// TwinCAT 3 PLC project _49001_01_BSM_762_V01_000_ISCOtherm
// libraries:
//   Tc2_EtherCAT, * (Beckhoff Automation GmbH)
//   Tc2_IoFunctions, * (Beckhoff Automation GmbH)
//   Tc2_Math, * (Beckhoff Automation GmbH)
//   Tc2_MC2, * (Beckhoff Automation GmbH)
//   Tc2_NC, * (Beckhoff Automation GmbH)
//   Tc2_NCI, * (Beckhoff Automation GmbH)
//   Tc2_SerialCom, * (Beckhoff Automation GmbH)
//   Tc2_Standard, * (Beckhoff Automation GmbH)
//   Tc2_System, * (Beckhoff Automation GmbH)
//   Tc2_Utilities, * (Beckhoff Automation GmbH)
//   Tc3_Module, * (Beckhoff Automation GmbH)
//   Lib1,1.0.0.0,riex
// project tree:
//   Data types/Machine/BECKHOFF/ ST_BECKHOFFDRIVETOPLC.TcDUT, ST_BECKHOFFDRIVE_REF.TcDUT, ST_PLCTOBECKHOFFDRIVE.TcDUT
//   Data types/Machine/FORCE/ ST_FORCETOPLC.TcDUT, ST_FORCE_REF.TcDUT, ST_PLCTOFORCE.TcDUT
//   Data types/Machine/Group_0000 - General/ ET_Gr00Auto.TcDUT, ET_Gr00Home.TcDUT, ST_Gr00HMIRef.TcDUT, ST_Gr00HMITOPLC.TcDUT, ST_Gr00PLCTOHMI.TcDUT
//   Data types/Machine/Group_0001/ ET_Gr01Auto.TcDUT, ET_Gr01Home.TcDUT, ET_Gr01HomeAxis.TcDUT, ET_Gr01HomeSawband.TcDUT, ET_Gr01Manual.TcDUT, ST_Gr01HMIRef.TcDUT, ST_Gr01HMITOPLC.TcDUT, ST_Gr01PLCTOHMI.TcDUT
//   Data types/Machine/Group_0002/ ET_Gr02Auto.TcDUT, ET_Gr02Home.TcDUT, ET_Gr02HomeAxis.TcDUT, ET_Gr02Manual.TcDUT, ST_Gr02HMIRef.TcDUT, ST_Gr02HMITOPLC.TcDUT, ST_Gr02PLCTOHMI.TcDUT
//   Data types/Machine/Group_0005/ ET_Gr05Auto.TcDUT, ET_Gr05AutoProcess.TcDUT, ET_Gr05Home.TcDUT, ET_Gr05HomeAxis.TcDUT, ET_Gr05HomeAxisClamp1.TcDUT, ET_Gr05Manual.TcDUT, ST_Gr05HMIRef.TcDUT, ST_Gr05HMITOPLC.TcDUT, ST_Gr05PLCTOHMI.TcDUT
//   Data types/Machine/SEW/CIA402/ ST_PLCTOSEWMOVIEDRIVEBCIA402.TcDUT, ST_SEWMOVIEDRIVEBCIA402TOPLC.TcDUT, ST_SEWMOVIEDRIVEBCIA402_REF.TcDUT
//   Data types/Machine/STOEBER/PS6A34/ ST_STOEBER_PS6A34Status.TcDUT
//   Data types/Machine/STOEBER/SDS/ ST_BaseDeviceIn.TcDUT, ST_BaseDeviceOut.TcDUT, ST_PLCTOSTOEBER.TcDUT, ST_STOEBERTOPLC.TcDUT
//   Data types/Machine/STOEBER/SI6_SC6/CIA402/ ST_CIA402In.TcDUT, ST_CIA402Out.TcDUT, ST_PLCTOSTOEBERSI6SC6CIA402.TcDUT, ST_STOEBERSI6SC6CIA402TOPLC.TcDUT, ST_STOEBERSI6SC6CIA402_REF.TcDUT
//   Data types/Machine/STOEBER/ ST_STOEBER_AxisStatus.TcDUT
//   Data types/Machine/WeldingPhases/ ET_WeldingDirection.TcDUT, ST_WeldingStatus.TcDUT
//   Data types/Machine/WeldingPhases/Force/ ST_BeadUp.TcDUT, ST_ForceProcess.TcDUT, ST_ForceWelding.TcDUT, ST_HeatUp.TcDUT, ST_PreHeat.TcDUT, ST_WeldingPhases.TcDUT
//   Data types/Machine/WeldingPhases/Position/ ST_PositionProcess.TcDUT, ST_PositionWelding.TcDUT
//   Data types/Objects/Axis/ExternelMC/ ET_JogMode.TcDUT, ET_MC_Direction.TcDUT, ET_MC_States.TcDUT, ST_AXIS_REF.TcDUT, ST_NCTOPLC.TcDUT, ST_PLCTONC.TcDUT
//   Data types/Objects/Axis/ExternelMC/SDS/ ST_CommandPositioningFROMNC.TcDUT, ST_CommandPositioningFROMPLC.TcDUT, ST_DRIVE_REF.TcDUT, ST_FastRefereneValueFROMNC.TcDUT, ST_FastRefereneValueFROMPLC.TcDUT
//   Data types/Objects/Axis/ExternelMC/SI6/ ET_ModesOfOperation.TcDUT, ST_DRIVESI6SC6CIA402_REF.TcDUT, ST_HomingModeFromDrive.TcDUT, ST_HomingModeFromPLC.TcDUT, ST_JogModeFromPLC.TcDUT, ST_PositionModeFromDrive.TcDUT, ST_PositionModeFromPLC.TcDUT, ST_TorqueModeFromDrive.TcDUT, ST_TorqueModeFromPLC.TcDUT, ST_VelocityModeFromDrive.TcDUT, ST_VelocityModeFromPLC.TcDUT
//   Data types/Objects/Axis/InternalMC/Controller/ ET_MC_ControllerMode.TcDUT, ST_VeloControllerConfig.TcDUT
//   Data types/Objects/Axis/InternalMC/Drive/Control/ ST_AxisCtrl.TcDUT (not stored), ST_TippingMode.TcDUT (not stored)
//   Data types/Objects/Axis/InternalMC/Drive/Parameter/ ST_Dynamics.TcDUT (not stored), ST_LimitSwitches.TcDUT (not stored), ST_Position.TcDUT (not stored)
//   Data types/Objects/Axis/InternalMC/Drive/Scaling/ ET_MC_RampType.TcDUT (not stored), ET_ScalingMethod.TcDUT (not stored), ST_Scaling.TcDUT (not stored)
//   Data types/Objects/Axis/InternalMC/Drive/States/ ET_MC_MotionStates.TcDUT (not stored), ST_AxisStates.TcDUT (not stored)
//   Data types/Objects/Axis/InternalMC/Drive/ ST_DriveConfig.TcDUT
//   Data types/Objects/Axis/InternalMC/Encoder/ ST_EncoderConfig.TcDUT
//   Data types/Objects/Axis/InternalMC/ ST_AXIS_REF_V2.TcDUT
//   Data types/Objects/EtherCAT Diag/ ET_EtherCATDiag.TcDUT, E_EcCommState.TcDUT, ST_EcMasterDevState.TcDUT, ST_SlaveState.TcDUT, ST_SlaveStateInfo.TcDUT, ST_SlaveStateInfoScanned.TcDUT, ST_TopologyData.TcDUT
//   Data types/Objects/ET_SpindleCtrl/ ET_SpindleCtrl.TcDUT
//   Data types/Objects/FB_Alarm/ ET_AlarmType.TcDUT, ST_Alarm.TcDUT, ST_AlarmIn.TcDUT, ST_AlarmOut.TcDUT, ST_AlarmProperties.TcDUT, ST_AlarmRef.TcDUT
//   Data types/Objects/FB_AxisController/ ET_AxisGetLimits.TcDUT, ET_AxisSetLimits.TcDUT, ET_STOEBER_AxisGetLimitsTc2.TcDUT, ET_STOEBER_AxisSetLimitsTc2.TcDUT
//   Data types/Objects/FB_AxisMoveManual/ ET_AxisMoveManualSetLimits.TcDUT
//   Data types/Objects/FB_Blinker/ ST_Blinker.TcDUT
//   Data types/Objects/FB_CalcContour/ ET_ContourType.TcDUT
//   Data types/Objects/FB_CfgAxisInExt3DGroup/ ET_CfgAxisInExt3DGroup.TcDUT
//   Data types/Objects/FB_DistanceCounter/ ST_DistanceCounter.TcDUT
//   Data types/Objects/FB_EL3312/ ET_EL3312ThermocoupleTyp.TcDUT, ST_EL3312ChannelState.TcDUT, ST_EL3312CoeInfo.TcDUT, ST_EL3312CoeReadData.TcDUT, ST_EL3312CoeWriteData.TcDUT
//   Data types/Objects/FB_EL3351/ ST_EL3351ChannelState.TcDUT, ST_EL3351CoeInfo.TcDUT, ST_EL3351CoeReadData.TcDUT, ST_EL3351CoeWriteData.TcDUT
//   Data types/Objects/FB_EL3356/ ST_EL3356ChannelCtrl.TcDUT, ST_EL3356ChannelState.TcDUT, ST_EL3356CoeInfo.TcDUT, ST_EL3356CoeReadData.TcDUT, ST_EL3356CoeWriteData.TcDUT
//   Data types/Objects/FB_ExtSetPoint/ ET_MoveExtState.TcDUT
//   Data types/Objects/FB_ExtTrajPos/ ET_CalcExtTrajState.TcDUT
//   Data types/Objects/FB_ItpReadRParams/ ET_ItpReadRParams.TcDUT
//   Data types/Objects/FB_ItpWriteRParams/ ET_ItpWriteRParams.TcDUT
//   Data types/Objects/FB_KL600x/ ET_KL600xInit.TcDUT, ET_KL600xSend.TcDUT, ST_KL600xData.TcDUT
//   Data types/Objects/FB_LoadFromFile/ ET_LoadFromFile.TcDUT
//   Data types/Objects/FB_Logger/ ST_Logger.TcDUT, ST_LoggerVar.TcDUT
//   Data types/Objects/FB_ModeSelector/ ET_MachineMode.TcDUT, ET_MachineState.TcDUT
//   Data types/Objects/FB_RampDirector/ ET_RampGenerator.TcDUT
//   Data types/Objects/FB_SpindlePreheat/ ET_SpindlePreheat.TcDUT, ST_SpindlePreheat.TcDUT
//   Data types/Objects/FB_TimeHoursCounter/ ST_TimeHoursCounter.TcDUT
//   Data types/Objects/FB_Timer/ ST_DateTime.TcDUT, ST_Time.TcDUT
//   Data types/Objects/FB_ToolStorage/ ET_ToolStatus.TcDUT, ET_ToolStorage.TcDUT
//   Data types/Objects/FB_Traceability/ ST_Traceability.TcDUT, ST_TraceabilityData.TcDUT, ST_TraceabilitySettings.TcDUT
//   Data types/Objects/Fieldbus/ ST_FieldbusStatus.TcDUT
//   Data types/Objects/Gefran/ ET_GFX4IR.TcDUT, ST_GFX4IRTOPLC.TcDUT, ST_GFX4IR_REF.TcDUT, ST_PLCTOGFX4IR.TcDUT
//   Data types/Objects/Leister/ ET_LeisterExtruder.TcDUT, ET_LeisterHeater.TcDUT, ST_LEISTERTOPLC.TcDUT, ST_LEISTER_REF.TcDUT, ST_PLCTOLEISTER.TcDUT
//   Data types/Objects/Munsch/ ET_MunschExtruder.TcDUT, ET_MUNSCH_CMD.TcDUT, ET_MUNSCH_RES.TcDUT, ST_MUNSCH_CMD_Data.TcDUT, ST_MUNSCH_REF.TcDUT, ST_MUNSCH_RES_Data.TcDUT
//   Data types/Objects/Periphery/ ST_PERIPHERYTOPLC.TcDUT, ST_PERIPHERY_REF.TcDUT, ST_PLCTOPERIPHERY.TcDUT
//   Data types/Objects/Robot/KUKA/ ET_KukaStart.TcDUT, ST_KUKATOPLC.TcDUT, ST_KUKA_REF.TcDUT, ST_PLCTOKUKA.TcDUT
//   Data types/Objects/Robot/ ST_PLCTOROBOT.TcDUT, ST_ROBOTTOPLC.TcDUT
//   Data types/Objects/Robot/YASKAWA/ ET_YaskawaStart.TcDUT, ST_PLCTOYASKAWA.TcDUT, ST_YASKAWATOPLC.TcDUT, ST_YASKAWA_REF.TcDUT
//   Data types/Objects/Spindle/ ET_SpindleClutchStatus.TcDUT
//   Data types/Objects/Spindle/PDS/ ST_SpindlePDSXLA170ClutchStatus.TcDUT, ST_SpindlePDSXLHClutchStatus.TcDUT
//   Data types/Objects/Terminal/ ST_TerminalState.TcDUT
//   Data types/Objects/TouchProbe/Renishaw/ ST_TouchProbeRenishawCtrl.TcDUT, ST_TouchProbeRenishawStatus.TcDUT
//   Data types/Objects/VFD/ ST_PLCTOVFD.TcDUT, ST_VFDTOPLC.TcDUT, ST_VFD_AXIS_REF.TcDUT, ST_VFD_DRIVE_REF.TcDUT
//   Global Variables/Alarms/ GVL_Gr00Alarm.TcGVL, GVL_Gr01Alarm.TcGVL, GVL_Gr02Alarm.TcGVL, GVL_Gr05Alarm.TcGVL
//   Global Variables/Basics/ GVL_FB_CheckArrayBounds.TcGVL, GVL_FB_CheckDivRealInfo.TcGVL
//   Global Variables/Config/ GVL_Gr00Config.TcGVL, GVL_Gr01Config.TcGVL, GVL_Gr02Config.TcGVL, GVL_Gr05Config.TcGVL
//   Global Variables/FB_Alarm/ GVL_FB_Alarm.TcGVL
//   Global Variables/FB_Fieldbus/ GVL_FB_Fieldbus.TcGVL
//   Global Variables/FB_GFX4IRZones/ GVL_FB_GFX4IRZones.TcGVL
//   Global Variables/FB_LoadFromFile/ GVL_FB_LoadFromFile.TcGVL
//   Global Variables/FB_Logger/ GVL_FB_Logger.TcGVL
//   Global Variables/FB_Traceability/ GVL_Traceability.TcGVL
//   Global Variables/ GVL.TcGVL, GVL_Gr0000.TcGVL, GVL_Gr0100.TcGVL, GVL_Gr0200.TcGVL, GVL_Gr0500.TcGVL, TwinCAT_Import.TcGVL
//   Global Variables/HMI/ GVL_Gr00HMI.TcGVL, GVL_Gr01HMI.TcGVL, GVL_Gr02HMI.TcGVL, GVL_Gr05HMI.TcGVL
//   Global Variables/Init/ GVL_Gr00Init.TcGVL, GVL_Gr01Init.TcGVL, GVL_Gr02Init.TcGVL, GVL_Gr05Init.TcGVL
//   Global Variables/Interface/ GVL_Gr00Interface.TcGVL, GVL_Gr01Interface.TcGVL, GVL_Gr02Interface.TcGVL, GVL_Gr05Interface.TcGVL
//   Global Variables/IO/ GVL_Gr00IO.TcGVL, GVL_Gr01IO.TcGVL, GVL_Gr02IO.TcGVL, GVL_Gr05IO.TcGVL
//   / PLC_TASK.TcTTO, Recipe Manager.TcRMO (not stored) (excluded from build)
//   POUs/ FAST.TcPOU, Init.TcPOU, MAIN.TcPOU
//   POUs/Machine/Group_0000 - General/Gr00Alarm/ FB_Gr00Alarm.TcPOU
//   POUs/Machine/Group_0000 - General/Gr00Control/ Gr00Control.TcPOU
//   POUs/Machine/Group_0000 - General/Gr00Control/Gr00Periphery/ FB_Gr00Periphery.TcPOU
//   POUs/Machine/Group_0000 - General/Gr00Control/Gr00Program/ FB_Gr00Program.TcPOU
//   POUs/Machine/Group_0000 - General/Gr00Control/Gr00Safety/ FB_Gr00Safety.TcPOU
//   POUs/Machine/Group_0000 - General/Gr00Control/Gr00Signals/ FB_Gr00Signals.TcPOU
//   POUs/Machine/Group_0000 - General/Gr00Control/Gr00Utility/ FB_Gr00Utility.TcPOU
//   POUs/Machine/Group_0000 - General/ Gr00Coordinator.TcPOU
//   POUs/Machine/Group_0000 - General/Gr00MachineMode/Gr00Auto/ Gr00Auto.TcPOU
//   POUs/Machine/Group_0000 - General/Gr00MachineMode/Gr00Auto/Gr00AutoAlarm/ FB_Gr00AutoAlarm.TcPOU (not stored)
//   POUs/Machine/Group_0000 - General/Gr00MachineMode/Gr00Auto/Gr00AutoInit/ FB_Gr00AutoInit.TcPOU (not stored)
//   POUs/Machine/Group_0000 - General/Gr00MachineMode/Gr00Auto/Gr00AutoProcedure/ FB_Gr00AutoProcedure.TcPOU (not stored)
//   POUs/Machine/Group_0000 - General/Gr00MachineMode/Gr00HMI/ Gr00HMI.TcPOU
//   POUs/Machine/Group_0000 - General/Gr00MachineMode/Gr00Home/ Gr00Home.TcPOU
//   POUs/Machine/Group_0000 - General/Gr00MachineMode/Gr00Home/Gr00HomeAlarm/ FB_Gr00HomeAlarm.TcPOU (not stored)
//   POUs/Machine/Group_0000 - General/Gr00MachineMode/Gr00Home/Gr00HomeInit/ FB_Gr00HomeInit.TcPOU (not stored)
//   POUs/Machine/Group_0000 - General/Gr00MachineMode/Gr00Home/Gr00HomeProcedure/ FB_Gr00HomeProcedure.TcPOU (not stored)
//   POUs/Machine/Group_0000 - General/Gr00MachineMode/ Gr00MachineMode.TcPOU
//   POUs/Machine/Group_0000 - General/Gr00MachineMode/Gr00Manual/ Gr00Manual.TcPOU
//   POUs/Machine/Group_0000 - General/Gr00MachineMode/Gr00Manual/Gr00ManualAlarm/ FB_Gr00ManualAlarm.TcPOU (not stored)
//   POUs/Machine/Group_0000 - General/Gr00MachineMode/Gr00Manual/Gr00ManualInit/ FB_Gr00ManualInit.TcPOU (not stored)
//   POUs/Machine/Group_0000 - General/Gr00MachineMode/Gr00Manual/Gr00ManualProcedure/ FB_Gr00ManualProcedure.TcPOU (not stored)
//   POUs/Machine/Group_0000 - General/Gr00Persistent/ Gr00Persistent.TcPOU
//   POUs/Machine/Group_0000 - General/Gr00Simulation/ Gr00Simulation.TcPOU
//   POUs/Machine/Group_0100 - Production/Gr01Control/Gr01Alarm/ FB_Gr01Alarm.TcPOU
//   POUs/Machine/Group_0100 - Production/Gr01Control/ Gr01Control.TcPOU
//   POUs/Machine/Group_0100 - Production/Gr01Control/Gr01Safety/ FB_Gr01Safety.TcPOU
//   POUs/Machine/Group_0100 - Production/Gr01Control/Gr01Signals/ FB_Gr01Signals.TcPOU
//   POUs/Machine/Group_0100 - Production/Gr01Control/Gr01Units/ FB_Gr01Angle.TcPOU, FB_Gr01SawBow.TcPOU
//   POUs/Machine/Group_0100 - Production/Gr01Control/Gr01Units/FB_Gr01Sawband/ FB_Gr01Sawband.TcPOU (not stored), FB_LowPassFilter.TcPOU (not stored), FB_PosVeloEnc.TcPOU (not stored)
//   POUs/Machine/Group_0100 - Production/Gr01Control/Gr01Utility/ FB_Gr01Utility.TcPOU
//   POUs/Machine/Group_0100 - Production/ Gr01Coordinator.TcPOU
//   POUs/Machine/Group_0100 - Production/Gr01HMI/ Gr01HMI.TcPOU
//   POUs/Machine/Group_0100 - Production/Gr01MachineMode/Gr01Auto/ Gr01Auto.TcPOU
//   POUs/Machine/Group_0100 - Production/Gr01MachineMode/Gr01Auto/Gr01AutoAlarm/ FB_Gr01AutoAlarm.TcPOU (not stored)
//   POUs/Machine/Group_0100 - Production/Gr01MachineMode/Gr01Auto/Gr01AutoInit/ FB_Gr01AutoInit.TcPOU (not stored)
//   POUs/Machine/Group_0100 - Production/Gr01MachineMode/Gr01Auto/Gr01AutoProcedure/ FB_Gr01AutoProcedure.TcPOU (not stored)
//   POUs/Machine/Group_0100 - Production/Gr01MachineMode/Gr01Home/ Gr01Home.TcPOU
//   POUs/Machine/Group_0100 - Production/Gr01MachineMode/Gr01Home/Gr01HomeAlarm/ FB_Gr01HomeAlarm.TcPOU (not stored)
//   POUs/Machine/Group_0100 - Production/Gr01MachineMode/Gr01Home/Gr01HomeFunctions/ FB_Gr01HomeAngle.TcPOU (not stored), FB_Gr01HomeAxisSawBow.TcPOU (not stored), FB_Gr01HomeSawband.TcPOU (not stored)
//   POUs/Machine/Group_0100 - Production/Gr01MachineMode/Gr01Home/Gr01HomeInit/ FB_Gr01HomeInit.TcPOU (not stored)
//   POUs/Machine/Group_0100 - Production/Gr01MachineMode/Gr01Home/Gr01HomeProcedure/ FB_Gr01HomeProcedure.TcPOU (not stored)
//   POUs/Machine/Group_0100 - Production/Gr01MachineMode/ Gr01MachineMode.TcPOU
//   POUs/Machine/Group_0100 - Production/Gr01MachineMode/Gr01Manual/ Gr01Manual.TcPOU
//   POUs/Machine/Group_0100 - Production/Gr01MachineMode/Gr01Manual/Gr01ManualAlarm/ FB_Gr01ManualAlarm.TcPOU (not stored)
//   POUs/Machine/Group_0100 - Production/Gr01MachineMode/Gr01Manual/Gr01ManualInit/ FB_Gr01ManualInit.TcPOU (not stored)
//   POUs/Machine/Group_0100 - Production/Gr01MachineMode/Gr01Manual/Gr01ManualProcedure/ FB_Gr01ManualProcedure.TcPOU (not stored)
//   POUs/Machine/Group_0100 - Production/Gr01Persistent/ Gr01Persistent.TcPOU
//   POUs/Machine/Group_0100 - Production/Gr01Simulation/ Gr01Simulation.TcPOU
//   POUs/Machine/Group_0500 - Transport/Gr05Control/Gr05Alarm/ FB_Gr05Alarm.TcPOU
//   POUs/Machine/Group_0500 - Transport/Gr05Control/ Gr05Control.TcPOU
//   POUs/Machine/Group_0500 - Transport/Gr05Control/Gr05Safety/ FB_Gr05Safety.TcPOU
//   POUs/Machine/Group_0500 - Transport/Gr05Control/Gr05Signals/ FB_Gr05Signals.TcPOU
//   POUs/Machine/Group_0500 - Transport/Gr05Control/Gr05Units/ FB_Gr05AxisClamp.TcPOU, FB_Gr05CylinderClamp.TcPOU, FB_Gr05CylinderPos.TcPOU, FB_Gr05RemovalBand.TcPOU, FB_Gr05Slide.TcPOU
//   POUs/Machine/Group_0500 - Transport/Gr05Control/Gr05Utility/ FB_Gr05Utility.TcPOU
//   POUs/Machine/Group_0500 - Transport/ Gr05Coordinator.TcPOU
//   POUs/Machine/Group_0500 - Transport/Gr05HMI/ Gr05HMI.TcPOU
//   POUs/Machine/Group_0500 - Transport/Gr05MachineMode/Gr05Auto/ Gr05Auto.TcPOU
//   POUs/Machine/Group_0500 - Transport/Gr05MachineMode/Gr05Auto/Gr05AutoAlarm/ FB_Gr05AutoAlarm.TcPOU (not stored)
//   POUs/Machine/Group_0500 - Transport/Gr05MachineMode/Gr05Auto/Gr05AutoInit/ FB_Gr05AutoInit.TcPOU (not stored)
//   POUs/Machine/Group_0500 - Transport/Gr05MachineMode/Gr05Auto/Gr05AutoProcedure/ FB_Gr05AutoProcedure.TcPOU (not stored)
//   POUs/Machine/Group_0500 - Transport/Gr05MachineMode/Gr05Home/ Gr05Home.TcPOU
//   POUs/Machine/Group_0500 - Transport/Gr05MachineMode/Gr05Home/Gr05HomeAlarm/ FB_Gr05HomeAlarm.TcPOU (not stored)
//   POUs/Machine/Group_0500 - Transport/Gr05MachineMode/Gr05Home/Gr05HomeFunctions/ FB_Gr05HomeAxisClamp1.TcPOU (not stored), FB_Gr05HomeAxisClamp2.TcPOU (not stored)
//   POUs/Machine/Group_0500 - Transport/Gr05MachineMode/Gr05Home/Gr05HomeInit/ FB_Gr05HomeInit.TcPOU (not stored)
//   POUs/Machine/Group_0500 - Transport/Gr05MachineMode/Gr05Home/Gr05HomeProcedure/ FB_Gr05HomeProcedure.TcPOU (not stored)
//   POUs/Machine/Group_0500 - Transport/Gr05MachineMode/ Gr05MachineMode.TcPOU
//   POUs/Machine/Group_0500 - Transport/Gr05MachineMode/Gr05Manual/ Gr05Manual.TcPOU
//   POUs/Machine/Group_0500 - Transport/Gr05MachineMode/Gr05Manual/Gr05ManualAlarm/ FB_Gr05ManualAlarm.TcPOU (not stored)
//   POUs/Machine/Group_0500 - Transport/Gr05MachineMode/Gr05Manual/Gr05ManualInit/ FB_Gr05ManualInit.TcPOU (not stored)
//   POUs/Machine/Group_0500 - Transport/Gr05MachineMode/Gr05Manual/Gr05ManualProcedure/ FB_Gr05ManualProcedure.TcPOU (not stored)
//   POUs/Machine/Group_0500 - Transport/Gr05Persistent/ Gr05Persistent.TcPOU
//   POUs/Machine/Group_0500 - Transport/Gr05Simulation/ Gr05Simulation.TcPOU
//   POUs/Tc2 Objects/Alarm/ FB_Alarm.TcPOU, FB_Error.TcPOU, FB_FatalError.TcPOU, FB_Hint.TcPOU, FB_Message.TcPOU, FB_Warning.TcPOU
//   POUs/Tc2 Objects/Automation/Axis/Beckhoff/CommandPositioning/ FB_AxisController.TcPOU (not stored), FB_AxisMoveAuto.TcPOU (not stored), FB_AxisMoveManual.TcPOU (not stored)
//   POUs/Tc2 Objects/Automation/Axis/Beckhoff/ FB_AxisMcBeckhoff.TcPOU, FB_AxisMcBeckhoffSEWMoviDriveBVelo.TcPOU, FB_AxisMcBeckhoffStoeberSCI6.TcPOU, FB_BECKHOFFDRIVE_REF.TcPOU
//   POUs/Tc2 Objects/Automation/Axis/ F_ChkAllAxisCoupled.TcPOU, F_ChkAllAxisEnabled.TcPOU, F_ChkAllAxisFieldbusOK.TcPOU, F_ChkAllAxisInSamePos.TcPOU, F_ChkAllAxisNotMoving.TcPOU, F_ChkAllAxisReferenced.TcPOU, F_ChkAllAxisStandStill.TcPOU
//   POUs/Tc2 Objects/Automation/Axis/OnOff/ FB_OnOff_AxisController.TcPOU, FB_OnOff_AxisMoveAuto.TcPOU, FB_OnOff_AxisMoveManual.TcPOU
//   POUs/Tc2 Objects/Automation/Axis/OnOff/Motion/ FB_OnOff_MoveAbsolut.TcPOU (not stored), FB_OnOff_MoveVelocity.TcPOU (not stored), FB_OnOff_Power.TcPOU (not stored), FB_OnOff_Reset.TcPOU (not stored), FB_OnOff_Stop.TcPOU (not stored)
//   POUs/Tc2 Objects/Automation/Axis/Override/ FB_Override.TcPOU, FB_OverrideSelection.TcPOU
//   POUs/Tc2 Objects/Automation/Axis/Own/Interface/Drive/ FB_AXIS_REF_V2.TcPOU (not stored)
//   POUs/Tc2 Objects/Automation/Axis/SEW/MOVIDRIVE B/ FB_SEWMOVIDRIVEBCIA402_REF.TcPOU (not stored)
//   POUs/Tc2 Objects/Automation/Axis/Stöber/SDS/CommandPositioning/ FB_AxisMcStoeber.TcPOU (not stored), FB_STOEBERSDS_MC_AxisController.TcPOU (not stored), FB_STOEBERSDS_MC_AxisMoveAuto.TcPOU (not stored), FB_STOEBERSDS_MC_AxisMoveManual.TcPOU (not stored), FB_STOEBERSDS_MC_GearIn.TcPOU (not stored), FB_STOEBERSDS_MC_GearOut.TcPOU (not stored), FB_STOEBERSDS_MC_Halt_noready.TcPOU (not stored), FB_STOEBERSDS_MC_Home.TcPOU (not stored), FB_STOEBERSDS_MC_Jog.TcPOU (not stored), FB_STOEBERSDS_MC_MoveAbsolut.TcPOU (not stored), FB_STOEBERSDS_MC_MoveAdditive.TcPOU (not stored), FB_STOEBERSDS_MC_MoveRelative.TcPOU (not stored), FB_STOEBERSDS_MC_MoveSuperimposed.TcPOU (not stored), FB_STOEBERSDS_MC_MoveVelocity.TcPOU (not stored), FB_STOEBERSDS_MC_Power.TcPOU (not stored), FB_STOEBERSDS_MC_Reset.TcPOU (not stored), FB_STOEBERSDS_MC_Stop.TcPOU (not stored), F_MoveToAxisRef.TcPOU (not stored)
//   POUs/Tc2 Objects/Automation/Axis/Stöber/SDS/FastRefereneValue/ FB_AxisStoeberSDS.TcPOU (not stored), FB_STOEBERSDS_AxisController.TcPOU (not stored), FB_STOEBERSDS_AxisMoveAuto.TcPOU (not stored), FB_STOEBERSDS_AxisMoveManual.TcPOU (not stored), FB_STOEBERSDS_Drive_REF.TcPOU (not stored), FB_STOEBERSDS_Home.TcPOU (not stored), FB_STOEBERSDS_Jog.TcPOU (not stored), FB_STOEBERSDS_MoveAbsolut.TcPOU (not stored), FB_STOEBERSDS_MoveVelocity.TcPOU (not stored), FB_STOEBERSDS_Power.TcPOU (not stored), FB_STOEBERSDS_QuickStop.TcPOU (not stored), FB_STOEBERSDS_Reset.TcPOU (not stored), FB_STOEBERSDS_Stop.TcPOU (not stored)
//   POUs/Tc2 Objects/Automation/Axis/Stöber/SDS/ FB_STOEBERSDS_AxisLink.TcPOU (not stored), FB_STOEBERSDS_ReadStatus.TcPOU (not stored)
//   POUs/Tc2 Objects/Automation/Axis/Stöber/SI6_SC6/ FB_StoeberPS6A34.TcPOU (not stored)
//   POUs/Tc2 Objects/Automation/Axis/VFD/ FB_VFD_AxisController.TcPOU, FB_VFD_AxisLink.TcPOU, FB_VFD_AxisMoveAuto.TcPOU, FB_VFD_AxisMoveManual.TcPOU (not stored), FB_VFD_Axis_REF.TcPOU (not stored), FB_VFD_Drive_REF.TcPOU (not stored), FB_VFD_MoveVelocity.TcPOU (not stored), FB_VFD_Power.TcPOU (not stored), FB_VFD_Reset.TcPOU (not stored), FB_VFD_Stop.TcPOU (not stored)
//   POUs/Tc2 Objects/Automation/Cylinder/ FB_Cylinder.TcPOU
//   POUs/Tc2 Objects/Automation/Cylinder/Hydraulic/ FB_HydraulicCylinder.TcPOU (not stored)
//   POUs/Tc2 Objects/Automation/Cylinder/Pneumatic/ FB_PneumaticCylinder.TcPOU (not stored)
//   POUs/Tc2 Objects/Automation/Cylinder/Position Cylinder/ FB_CylinderPos.TcPOU (not stored), FB_CylinderPos_MoveAbsolut.TcPOU (not stored), F_GetCylinderPos.TcPOU (not stored), F_SetCylinderPos.TcPOU (not stored)
//   POUs/Tc2 Objects/Automation/Extraction Fan/ FB_ExtractionFan.TcPOU
//   POUs/Tc2 Objects/Automation/Force/ FB_ForceController.TcPOU, FB_ForceReg.TcPOU, FB_FORCE_REF.TcPOU, FB_PID_Regler.TcPOU
//   POUs/Tc2 Objects/Automation/Heater/ FB_Heater.TcPOU
//   POUs/Tc2 Objects/Automation/MotorOnOff/ FB_Motor.TcPOU
//   POUs/Tc2 Objects/Automation/NCiChannel/ FB_CfgAxisInExt3DGroup.TcPOU
//   POUs/Tc2 Objects/Automation/NCiChannel/R-parameters/ FB_ItpReadRParams.TcPOU (not stored), FB_ItpWriteRParams.TcPOU (not stored)
//   POUs/Tc2 Objects/Automation/OperationMode/ FB_ModeSelector.TcPOU
//   POUs/Tc2 Objects/Automation/Process/ FB_StartProcess.TcPOU
//   POUs/Tc2 Objects/Automation/Sawband/ FB_Sawband.TcPOU
//   POUs/Tc2 Objects/Automation/Spindle/ FB_CoolingDevice.TcPOU, FB_SpindlePreheat.TcPOU, FB_ToolStorage.TcPOU, FB_VFD_SpindlePreheat.TcPOU, F_SpindleHSDClutchStatus.TcPOU, F_SpindlePDSXLA170ClutchStatus.TcPOU, F_SpindlePDSXLHClutchStatus.TcPOU
//   POUs/Tc2 Objects/Automation/Vacuum/ FB_Vacuum.TcPOU
//   POUs/Tc2 Objects/Basics/ CheckBounds.TcPOU (excluded from build), CheckDivReal.TcPOU (excluded from build), FB_CheckArrayBounds.TcPOU (excluded from build), FB_CheckDivRealInfo.TcPOU (excluded from build), FB_Get_Time.TcPOU, F_AdsError_Text.TcPOU
//   POUs/Tc2 Objects/Conversions/BitOriented/ F_ConvArrBitsToWord.TcPOU
//   POUs/Tc2 Objects/Diagnostic/Terminal/ FB_TerminalDiagnosis.TcPOU, FB_ToggleBit.TcPOU, F_StateReturn.TcPOU
//   POUs/Tc2 Objects/Engineering/Buffer/ FB_FiFo.TcPOU
//   POUs/Tc2 Objects/Engineering/Dynamics/CalcVeloAccDecJerk/ FB_CalcVeloAccDecJerk.TcPOU (not stored)
//   POUs/Tc2 Objects/Engineering/External set value generator/ FB_ExtSetPoint.TcPOU
//   POUs/Tc2 Objects/Engineering/Filter/ FB_PT1.TcPOU, FB_ValueFilter.TcPOU
//   POUs/Tc2 Objects/Engineering/Position offset/ F_PosOffset.TcPOU
//   POUs/Tc2 Objects/Engineering/Position/Controller/PID Components/ FB_CompD.TcPOU (not stored), FB_CompI.TcPOU (not stored), FB_CompP.TcPOU (not stored)
//   POUs/Tc2 Objects/Engineering/Position/Controller/PID Controller/ FB_CtrlOut.TcPOU (not stored), FB_CtrlPI.TcPOU (not stored), FB_CtrlPID.TcPOU (not stored), F_CtrlIn.TcPOU (not stored)
//   POUs/Tc2 Objects/Engineering/Position/Controller/PID Types/ FB_TypePI.TcPOU (not stored), FB_TypePID.TcPOU (not stored), FB_TypePIDW.TcPOU (not stored), FB_TypePIW.TcPOU (not stored)
//   POUs/Tc2 Objects/Engineering/Position/Controller/PositionController/ FB_PosCtrlIn.TcPOU (not stored), FB_PosCtrlOut.TcPOU (not stored), FB_PositionController.TcPOU (not stored)
//   POUs/Tc2 Objects/Engineering/Position/Encoder/ FB_PositionEncoder.TcPOU (not stored)
//   POUs/Tc2 Objects/Engineering/Position/ F_ModuloDistance.TcPOU
//   POUs/Tc2 Objects/Engineering/Position/Residuals/ F_ConvertActPosResiduals.TcPOU (not stored), F_ConvertSetPosResiduals.TcPOU (not stored)
//   POUs/Tc2 Objects/Engineering/Trajectory model/ FB_ExtContour.TcPOU, FB_ExtTraj.TcPOU, F_CalcContour.TcPOU, F_CalcTrajPos.TcPOU
//   POUs/Tc2 Objects/ExternalHardware/Beckhoff/EL..KL600x/ FB_KL600xData.TcPOU (not stored), FB_KL600xString.TcPOU (not stored)
//   POUs/Tc2 Objects/ExternalHardware/Beckhoff/EL3312/ FB_EL3312.TcPOU (not stored), FB_EL3312ChannelDiagnosis.TcPOU (not stored), FB_EL3312CoE.TcPOU (not stored)
//   POUs/Tc2 Objects/ExternalHardware/Beckhoff/EL3351/ FB_EL3351.TcPOU (not stored), FB_EL3351ChannelDiagnosis.TcPOU (not stored), FB_EL3351CoE.TcPOU (not stored), FB_EL3351Measuring.TcPOU (not stored)
//   POUs/Tc2 Objects/ExternalHardware/Beckhoff/EL3356/ FB_EL3356.TcPOU (not stored), FB_EL3356ChannelDiagnosis.TcPOU (not stored), FB_EL3356CoE.TcPOU (not stored)
//   POUs/Tc2 Objects/ExternalHardware/Gefran/ FB_GFX4IRCtrlZone.TcPOU, FB_GFX4IRZones.TcPOU, FB_GFX4IR_REF.TcPOU, F_ChkAllZonesNotEnabled.TcPOU
//   POUs/Tc2 Objects/ExternalHardware/KUKA/ FB_KUKA_Enable.TcPOU, FB_KUKA_Power.TcPOU, FB_KUKA_Prg.TcPOU, FB_KUKA_REF.TcPOU, FB_KUKA_Reset.TcPOU, FB_KUKA_StartProg.TcPOU, FB_MoveToKukaRef.TcPOU
//   POUs/Tc2 Objects/ExternalHardware/Leister/ FB_LeisterExtruder_Extruder.TcPOU, FB_LeisterExtruder_Heater.TcPOU, FB_LEISTER_EXTRUDER_REF.TcPOU
//   POUs/Tc2 Objects/ExternalHardware/Munsch/ FB_MunschExtruder.TcPOU, FB_MunschExtruderAir.TcPOU, FB_MunschExtruder_AirTemp.TcPOU, FB_MunschExtruder_Extruding.TcPOU, FB_MunschExtruder_Heat.TcPOU, FB_MunschExtruder_MaterialTemp.TcPOU, FB_MunschExtruder_ReadStatus.TcPOU, FB_MUNSCH_EXTRUDER_REF.TcPOU, F_MunschCMD.TcPOU, F_MunschRES.TcPOU
//   POUs/Tc2 Objects/ExternalHardware/Periphery/ FB_PERIPHERY_REF.TcPOU
//   POUs/Tc2 Objects/ExternalHardware/YASKAWA/ FB_YASKAWA_Controller.TcPOU, FB_YASKAWA_Power.TcPOU, FB_YASKAWA_REF.TcPOU, FB_YASKAWA_Reset.TcPOU, FB_YASKAWA_StartPrg.TcPOU
//   POUs/Tc2 Objects/File/ FB_FileHandler.TcPOU, FB_FileHandlerBinary.TcPOU, FB_LoadFromFile.TcPOU
//   POUs/Tc2 Objects/Logger/ FB_Logger.TcPOU, FB_LoggerFile.TcPOU
//   POUs/Tc2 Objects/Logic/ F_DwordToBitReal.TcPOU, F_RealToBitDword.TcPOU, F_ResetBitOfDWord.TcPOU, F_SetBitOfDWord.TcPOU
//   POUs/Tc2 Objects/Logic/Oscat/ CHECK_PARITY.TcPOU
//   POUs/Tc2 Objects/MachineEquipment/ F_AxisClamp2Pos.TcPOU, F_kAngleActuatorSpeedLin.TcPOU, F_kFeedReductionSlowGuidings.TcPOU
//   POUs/Tc2 Objects/Mathematical/Delay/ FB_Delay.TcPOU
//   POUs/Tc2 Objects/Mathematical/ FB_Differential.TcPOU, FB_Integral.TcPOU, F_Exp10.TcPOU, F_FloorDN.TcPOU, F_FracR.TcPOU, F_GCD.TcPOU, F_LRealRound.TcPOU, F_MM_TO_DEG.TcPOU, F_ModDW.TcPOU, F_ModR.TcPOU, F_RoundR.TcPOU
//   POUs/Tc2 Objects/Mathematical/Hysteresis/ FB_Hysteresis.TcPOU
//   POUs/Tc2 Objects/Mathematical/Limits/ FB_Limiter.TcPOU, F_DeadZone.TcPOU, F_WordToRange.TcPOU
//   POUs/Tc2 Objects/Mathematical/Scaling/ FB_Scaling.TcPOU, FB_ScalingOffset.TcPOU
//   POUs/Tc2 Objects/Measurements/Counter/ FB_Counter.TcPOU, FB_DistanceCounter.TcPOU, FB_TimeHoursCounter.TcPOU
//   POUs/Tc2 Objects/Measurements/ FB_TemperaturOK.TcPOU, FB_Timer.TcPOU
//   POUs/Tc2 Objects/Measurements/Oscat/ T_PLC_MS.TcPOU
//   POUs/Tc2 Objects/Measurements/RTC/ FB_RTC.TcPOU
//   POUs/Tc2 Objects/Safety/ FB_AirPressure.TcPOU, FB_LightCurtain.TcPOU, FB_NoEmergencyStop.TcPOU, FB_PowerSupply.TcPOU, FB_Temperature.TcPOU
//   POUs/Tc2 Objects/Safety/Fieldbus/ FB_EtherCATDiag.TcPOU, FB_EtherCATFrameDiag.TcPOU, FB_Fieldbus.TcPOU, FB_Fieldbus_v2.TcPOU
//   POUs/Tc2 Objects/Signals/Force Input/ FB_ForceBit.TcPOU, FB_ForceByte.TcPOU
//   POUs/Tc2 Objects/Signals/Generators/ FB_Blinker.TcPOU
//   POUs/Tc2 Objects/Signals/Handling/ FB_SignalHandlingDelay.TcPOU, FB_SignalHandlingEdge.TcPOU, F_SignalHandling.TcPOU
//   POUs/Tc2 Objects/Signals/Ramp Generators/ FB_RampDirector.TcPOU
//   POUs/Tc2 Objects/Signals/Ramp Generators/Oscat_Ramp/ FB_RMP_W.TcPOU (not stored), _RMP_W.TcPOU (not stored)
//   POUs/Tc2 Objects/Signals/Watchdog/ FB_SignalWatchdog.TcPOU, FB_SignalWatchdog2.TcPOU
//   POUs/Tc2 Objects/String/ F_CheckStringIsReal.TcPOU, F_RealToStrf.TcPOU
//   POUs/Tc2 Objects/Traceability/ FB_Traceability.TcPOU
//   POUs/Tc3 Objects/Alarm/ ET_AlarmType_1.TcDUT, FB_Alarm_1.TcPOU, FB_Error_1.TcPOU, FB_FatalError_1.TcPOU, FB_Hint_1.TcPOU, FB_Message_1.TcPOU, FB_Warning_1.TcPOU, GVL_FB_Alarm_1.TcGVL, ST_AlarmIn_1.TcDUT, ST_AlarmOut_1.TcDUT, ST_AlarmProperties_1.TcDUT, ST_AlarmRef_1.TcDUT, ST_Alarm_1.TcDUT
//   POUs/Tc3 Objects/Automation/Axis/Beckhoff/CommandPositioning/ ET_BECKHOFF_AxisGetLimits.TcDUT (not stored), ET_BECKHOFF_AxisSetLimits.TcDUT (not stored), ET_BECKHOFF_ManualSetLimits.TcDUT (not stored), FB_BECKHOFF_AxisController.TcPOU (not stored), FB_BECKHOFF_AxisMoveAuto.TcPOU (not stored), FB_BECKHOFF_AxisMoveManual.TcPOU (not stored)
//   POUs/Tc3 Objects/Automation/Axis/Bosch/CommandPositioning/Beckhoff/ ET_BOSCH_AxisGetLimits.TcDUT (not stored), ET_BOSCH_AxisSetLimits.TcDUT (not stored), ET_BOSCH_Home.TcDUT (not stored), ET_BOSCH_ManualSetLimits.TcDUT (not stored), ET_BOSCH_Reset.TcDUT (not stored), FB_AxisMcBeckhoffBoschIndraDrive.TcPOU (not stored), FB_BOSCH_AxisController.TcPOU (not stored), FB_BOSCH_AxisMoveAuto.TcPOU (not stored), FB_BOSCH_AxisMoveManual.TcPOU (not stored), FB_BOSCH_Home.TcPOU (not stored), FB_BOSCH_Reset.TcPOU (not stored)
//   POUs/Tc3 Objects/Automation/Axis/Bosch/Drive/ FB_BOSCH_DriveLink.TcPOU (not stored)
//   POUs/Tc3 Objects/Automation/Axis/Bosch/Drive/IndraDrive/ FB_BOSCHINDRADRIVECIA402_REF.TcPOU (not stored), ST_BOSCHINDRADRIVECIA402TOPLC.TcDUT (not stored), ST_BOSCHINDRADRIVECIA402_REF.TcDUT (not stored), ST_PLCTOBOSCHINDRADRIVECIA402.TcDUT (not stored)
//   POUs/Tc3 Objects/Automation/Axis/Bosch/ProcessController/ ET_BOSCH_ProcessCtrl.TcDUT (not stored), ET_BOSCH_ProcessCtrlGetValue.TcDUT (not stored), ET_BOSCH_ProcessCtrlSetValue.TcDUT (not stored), FB_BOSCH_ProcessCtrl.TcPOU (not stored), FB_BOSCH_ProcessCtrlLink.TcPOU (not stored), FB_BOSCH_ProcessCtrl_Reset.TcPOU (not stored), FB_BOSCH_ProcessCtrl_Start.TcPOU (not stored), FB_BOSCH_ProcessCtrl_Stop.TcPOU (not stored), ST_FWS_MLDPCx_PRE_01Vxx_MPxx.TcDUT (not stored)
//   POUs/Tc3 Objects/Automation/Axis/ F_ChkAllAxisCoupled_1.TcPOU, F_ChkAllAxisEnabled_1.TcPOU, F_ChkAllAxisInSamePos_1.TcPOU, F_ChkAllAxisNotMoving_1.TcPOU, F_ChkAllAxisReferenced_1.TcPOU, F_ChkAllAxisStandStill_1.TcPOU, F_ChkAxisError.TcPOU
//   POUs/Tc3 Objects/Automation/Axis/Stöber/CommandPositioning/Beckhoff/ ET_STOEBER_AxisGetLimits.TcDUT (not stored), ET_STOEBER_AxisSetLimits.TcDUT (not stored), ET_STOEBER_ManualSetLimits.TcDUT (not stored), FB_STOEBER_AxisController.TcPOU (not stored), FB_STOEBER_AxisMoveAuto.TcPOU (not stored), FB_STOEBER_AxisMoveManual.TcPOU (not stored)
//   POUs/Tc3 Objects/Automation/Axis/Stöber/Dirve/SI6SC6/ FB_STOEBERSI6SC6CIA402_REF.TcPOU (not stored), ST_PLCTOSTOEBERSI6SC6CIA402_1.TcDUT (not stored), ST_STOEBERSI6SC6CIA402TOPLC_1.TcDUT (not stored), ST_STOEBERSI6SC6CIA402_REF_1.TcDUT (not stored)
//   POUs/Tc3 Objects/Automation/Axis/Stöber/PS6A34/ ST_STOEBER_PS6A34Status_1.TcDUT (not stored)
//   POUs/Tc3 Objects/Automation/Cylinder/ FB_Cylinder_1.TcPOU
//   POUs/Tc3 Objects/Automation/Cylinder/Hydraulic/ FB_HydraulicCylinder_1.TcPOU (not stored)
//   POUs/Tc3 Objects/Automation/Cylinder/Pneumatic/ FB_PneumaticCylinder_1.TcPOU (not stored)
//   POUs/Tc3 Objects/Automation/Cylinder/Position Cylinder/ FB_PosCylinder.TcPOU (not stored), FB_PosCylinder_MoveAbsolut.TcPOU (not stored), F_GetPosCylinder.TcPOU (not stored), F_SetPosCylinder.TcPOU (not stored)
//   POUs/Tc3 Objects/Automation/Force/ FB_ForceController_1.TcPOU, FB_ForceReg_1.TcPOU, FB_PID_Regler_1.TcPOU
//   POUs/Tc3 Objects/Automation/NCiChannel/CfgAxisInExt3DGroup/ ET_CfgAxisInExt3DGroup_1.TcDUT (not stored), FB_CfgAxisInExt3DGroup_1.TcPOU (not stored)
//   POUs/Tc3 Objects/Automation/NCiChannel/ItpReadRParams/ ET_ItpReadRParams_1.TcDUT (not stored), FB_ItpReadRParams_1.TcPOU (not stored)
//   POUs/Tc3 Objects/Automation/NCiChannel/ItpWriteRParams/ ET_ItpWriteRParams_1.TcDUT (not stored), FB_ItpWriteRParams_1.TcPOU (not stored)
//   POUs/Tc3 Objects/Automation/OperationMode/ ET_MachineMode_1.TcDUT, ET_MachineState_1.TcDUT, ET_MaintenanceType.TcDUT, FB_ModeSelector_1.TcPOU
//   POUs/Tc3 Objects/Automation/Override/ FB_OverrideSelection_1.TcPOU, FB_Override_1.TcPOU
//   POUs/Tc3 Objects/Automation/Process/ FB_StartProcess_1.TcPOU
//   POUs/Tc3 Objects/Automation/Spindle/Clutch/ ET_SpindleClutchStatus_1.TcDUT (not stored), F_SpindleClutchStatus.TcPOU (not stored)
//   POUs/Tc3 Objects/Automation/Spindle/ FB_CoolingDevice_1.TcPOU
//   POUs/Tc3 Objects/Automation/Spindle/HSD/ F_SpindleHSDES951ClutchStatus.TcPOU (not stored), ST_SpindleHSDES951ClutchStatus.TcDUT (not stored)
//   POUs/Tc3 Objects/Automation/Spindle/PDS/ F_SpindlePDSXLA170ClutchStatus_1.TcPOU (not stored), ST_SpindlePDSXLA170ClutchStatus_1.TcDUT (not stored)
//   POUs/Tc3 Objects/Automation/Spindle/Preheat/ ET_SpindlePreheat_1.TcDUT (not stored), FB_SpindlePreheat_1.TcPOU (not stored), ST_SpindlePreheat_1.TcDUT (not stored)
//   POUs/Tc3 Objects/Automation/Vacuum/ FB_Vacuum_1.TcPOU
//   POUs/Tc3 Objects/Basics/ CheckBounds_1.TcPOU (excluded from build), CheckDivReal_1.TcPOU (excluded from build), FB_CheckArrayBounds_1.TcPOU (excluded from build), FB_CheckDivRealInfo_1.TcPOU (excluded from build), FB_Get_Time_1.TcPOU, F_AdsError_Text_1.TcPOU
//   POUs/Tc3 Objects/Communication/TCPIP/ASCII/ClientASCII/ FB_ClientASCIConnection.TcPOU (not stored), FB_ClientLogger.TcPOU (not stored), FB_ClientReceiveMsg.TcPOU (not stored), FB_ClientSendMsg.TcPOU (not stored)
//   POUs/Tc3 Objects/Communication/TCPIP/ ET_TCPIP_ConnectionState.TcDUT, GVL_TCPIP.TcGVL
//   POUs/Tc3 Objects/Communication/TCPIP/Helper/ FB_FrameFifo.TcPOU (not stored), FB_LogFifo.TcPOU (not stored)
//   POUs/Tc3 Objects/Conversions/BitOriented/ F_ConvArrBitsToWord_1.TcPOU
//   POUs/Tc3 Objects/Diagnostic/Terminal/ FB_TerminalDiagnosis_1.TcPOU, FB_ToggleBit_1.TcPOU, FUN_StateReturn.TcPOU, ST_TerminalState_1.TcDUT
//   POUs/Tc3 Objects/Engineering/Buffer/ FB_FiFo_1.TcPOU
//   POUs/Tc3 Objects/Engineering/Dynamics/CalcVeloAccDecJerk/ FB_CalcVeloAccDecJerk_1.TcPOU (not stored)
//   POUs/Tc3 Objects/Engineering/External set value generator/ ET_ExtSetpoint.TcDUT, FB_ExtSetpoint_1.TcPOU
//   POUs/Tc3 Objects/Engineering/Filter/ FB_PT1_1.TcPOU, FB_ValueFilter_1.TcPOU
//   POUs/Tc3 Objects/Engineering/Motion model/Contour/ ET_ContourType_1.TcDUT (not stored), FB_ExtContour_1.TcPOU (not stored), F_CalcContour_1.TcPOU (not stored)
//   POUs/Tc3 Objects/Engineering/Motion model/Oval/ ET_CalcExtOvalState.TcDUT (not stored), FB_ExtOval.TcPOU (not stored), F_CalcOval.TcPOU (not stored)
//   POUs/Tc3 Objects/Engineering/Motion model/Tilt/ ET_CalcExtTiltState.TcDUT (not stored), FB_ExtTilt.TcPOU (not stored), F_CalcTiltPos.TcPOU (not stored)
//   POUs/Tc3 Objects/Engineering/Motion model/Traj/ ET_CalcExtTrajState_1.TcDUT (not stored), FB_ExtTraj_1.TcPOU (not stored), F_CalcTrajPos_1.TcPOU (not stored)
//   POUs/Tc3 Objects/Engineering/Position offset/ F_PosOffset_1.TcPOU
//   POUs/Tc3 Objects/Engineering/Position/Controller/PID Components/ FB_CompD_1.TcPOU (not stored), FB_CompI_1.TcPOU (not stored), FB_CompP_1.TcPOU (not stored)
//   POUs/Tc3 Objects/Engineering/Position/Controller/PID CO_Ntroller/ FB_CtrlOut_1.TcPOU (not stored), FB_CtrlPID_1.TcPOU (not stored), FB_CtrlPI_1.TcPOU (not stored), F_CtrlIn_1.TcPOU (not stored)
//   POUs/Tc3 Objects/Engineering/Position/Controller/PID Types/ FB_TypePIDW_1.TcPOU (not stored), FB_TypePID_1.TcPOU (not stored), FB_TypePIW_1.TcPOU (not stored), FB_TypePI_1.TcPOU (not stored)
//   POUs/Tc3 Objects/Engineering/Position/Controller/PositionCO_Ntroller/ FB_PosCtrlIn_1.TcPOU (not stored), FB_PosCtrlOut_1.TcPOU (not stored), FB_PositionController_1.TcPOU (not stored)
//   POUs/Tc3 Objects/Engineering/Position/Encoder/ FB_PositionEncoder_1.TcPOU (not stored)
//   POUs/Tc3 Objects/Engineering/Position/ F_ModuloDistance_1.TcPOU
//   POUs/Tc3 Objects/Engineering/Position/Residuals/ F_ConvertActPosResiduals_1.TcPOU (not stored), F_ConvertSetPosResiduals_1.TcPOU (not stored)
//   POUs/Tc3 Objects/ExternalHardware/Beckhoff/EL..KL600x/ FB_KL600xData_1.TcPOU (not stored), FB_KL600xString_1.TcPOU (not stored)
//   POUs/Tc3 Objects/ExternalHardware/Beckhoff/EL3214/ ET_EL3214RTDElement.TcDUT (not stored), FB_EL3214.TcPOU (not stored), FB_EL3214ChannelDiagnosis.TcPOU (not stored), FB_EL3214CoE.TcPOU (not stored), ST_EL3214ChannelState.TcDUT (not stored), ST_EL3214CoeInfo.TcDUT (not stored), ST_EL3214CoeReadData.TcDUT (not stored), ST_EL3214CoeWriteData.TcDUT (not stored)
//   POUs/Tc3 Objects/ExternalHardware/Beckhoff/EL3312/ ET_EL3312ThermocoupleTyp_1.TcDUT (not stored), FB_EL3312ChannelDiagnosis_1.TcPOU (not stored), FB_EL3312CoE_1.TcPOU (not stored), FB_EL3312_1.TcPOU (not stored), ST_EL3312ChannelState_1.TcDUT (not stored), ST_EL3312CoeInfo_1.TcDUT (not stored), ST_EL3312CoeReadData_1.TcDUT (not stored), ST_EL3312CoeWriteData_1.TcDUT (not stored)
//   POUs/Tc3 Objects/ExternalHardware/Beckhoff/EL3351/ FB_EL3351ChannelDiagnosis_1.TcPOU (not stored), FB_EL3351CoE_1.TcPOU (not stored), FB_EL3351Measuring_1.TcPOU (not stored), FB_EL3351_1.TcPOU (not stored), ST_EL3351ChannelState_1.TcDUT (not stored), ST_EL3351CoeInfo_1.TcDUT (not stored), ST_EL3351CoeReadData_1.TcDUT (not stored), ST_EL3351CoeWriteData_1.TcDUT (not stored)
//   POUs/Tc3 Objects/ExternalHardware/Beckhoff/EL3356/ FB_EL3356ChannelDiagnosis_1.TcPOU (not stored), FB_EL3356CoE_1.TcPOU (not stored), FB_EL3356_1.TcPOU (not stored), ST_EL3356ChannelCtrl_1.TcDUT (not stored), ST_EL3356ChannelState_1.TcDUT (not stored), ST_EL3356CoeInfo_1.TcDUT (not stored), ST_EL3356CoeReadData_1.TcDUT (not stored), ST_EL3356CoeWriteData_1.TcDUT (not stored)
//   POUs/Tc3 Objects/ExternalHardware/Cognex/Scanner/ ET_COGNEX_ScannerCtrl.TcDUT (not stored), FB_DatamanScanner.TcPOU (not stored), FB_Scanner.TcPOU (not stored)
//   POUs/Tc3 Objects/ExternalHardware/Gefran/ ET_GFX4IR_1.TcDUT, FB_GFX4IRCtrlZone_1.TcPOU, FB_GFX4IRZones_1.TcPOU, FB_GFX4IR_REF_1.TcPOU, F_ChkAllZonesNotEnabled_1.TcPOU, GVL_GFX4IR.TcGVL, ST_GFX4IRTOPLC_1.TcDUT, ST_GFX4IR_REF_1.TcDUT, ST_PLCTOGFX4IR_1.TcDUT
//   POUs/Tc3 Objects/ExternalHardware/KUKA/ ET_KukaStart_1.TcDUT, FB_KUKA_Enable_1.TcPOU, FB_KUKA_Power_1.TcPOU, FB_KUKA_Prg_1.TcPOU, FB_KUKA_REF_1.TcPOU, FB_KUKA_Reset_1.TcPOU, FB_KUKA_StartProg_1.TcPOU, FB_MoveToKukaRef_1.TcPOU, ST_KUKATOPLC_1.TcDUT, ST_KUKA_REF_1.TcDUT, ST_PLCTOKUKA_1.TcDUT
//   POUs/Tc3 Objects/ExternalHardware/Munsch/ FB_MunschExtruderAir_1.TcPOU, FB_MunschExtruder_1.TcPOU, FB_MunschExtruder_AirTemp_1.TcPOU, FB_MunschExtruder_Heat_1.TcPOU, FB_MunschExtruder_MaterialTemp_1.TcPOU, FB_MunschExtruder_ReadStatus_1.TcPOU, FB_MUNSCH_EXTRUDER_REF_1.TcPOU, F_MunschCMD_1.TcPOU, F_MunschRES_1.TcPOU
//   POUs/Tc3 Objects/ExternalHardware/Periphery/ FB_PERIPHERY_REF_1.TcPOU, ST_PERIPHERY_REF_1.TcDUT, ST_PLC01TOPLC02.TcDUT, ST_PLC02TOPLC01.TcDUT, ST_PLC02TOPLC03.TcDUT, ST_PLC03TOPLC02.TcDUT
//   POUs/Tc3 Objects/ExternalHardware/Robot/ ST_PLCTOROBOT_1.TcDUT, ST_ROBOTTOPLC_1.TcDUT
//   POUs/Tc3 Objects/ExternalHardware/YASKAWA/ ET_YaskawaStart_1.TcDUT, FB_YASKAWA_Controller_1.TcPOU, FB_YASKAWA_Power_1.TcPOU, FB_YASKAWA_REF_1.TcPOU, FB_YASKAWA_Reset_1.TcPOU, FB_YASKAWA_StartPrg_1.TcPOU, ST_PLCTOYASKAWA_1.TcDUT, ST_YASKAWATOPLC_1.TcDUT, ST_YASKAWA_REF_1.TcDUT
//   POUs/Tc3 Objects/File/CSV/ ET_CSV_State.TcDUT, FB_FileCSVHandler.TcPOU, GVL_CSV.TcGVL
//   POUs/Tc3 Objects/File/TXT/ ET_LoadFromFile_1.TcDUT, FB_FileHandlerBinary_1.TcPOU, FB_FileHandler_1.TcPOU, FB_LoadFromFile_1.TcPOU, GVL_FB_LoadFromFile_1.TcGVL
//   POUs/Tc3 Objects/Logger/ FB_LoggerFile_1.TcPOU, FB_Logger_1.TcPOU, GVL_Logger.TcGVL, ST_LoggerVar_1.TcDUT, ST_Logger_1.TcDUT
//   POUs/Tc3 Objects/Logic/ F_DwordToBitReal_1.TcPOU, F_RealToBitDword_1.TcPOU, F_ResetBitOfDWord_1.TcPOU, F_SetBitOfDWord_1.TcPOU
//   POUs/Tc3 Objects/Logic/Oscat/ CHECK_PARITY_1.TcPOU
//   POUs/Tc3 Objects/Mathematical/Delay/ FB_Delay_1.TcPOU
//   POUs/Tc3 Objects/Mathematical/ FB_Differential_1.TcPOU, FB_Integral_1.TcPOU, F_Exp10_1.TcPOU, F_FloorDN_1.TcPOU, F_FracR_1.TcPOU, F_GCD_1.TcPOU, F_LRealRound_1.TcPOU, F_ModDW_1.TcPOU, F_ModR_1.TcPOU, F_RoundR_1.TcPOU
//   POUs/Tc3 Objects/Mathematical/Hysteresis/ FB_Hysteresis_1.TcPOU
//   POUs/Tc3 Objects/Mathematical/Limits/ FB_Limiter_1.TcPOU, F_DeadZone_1.TcPOU, F_WordToRange_1.TcPOU
//   POUs/Tc3 Objects/Mathematical/Scaling/ FB_ScalingOffset_1.TcPOU, FB_Scaling_1.TcPOU
//   POUs/Tc3 Objects/Measurements/Counter/ FB_Counter_1.TcPOU, FB_DistanceCounter_1.TcPOU, FB_TimeHoursCounter_1.TcPOU, ST_TimeHoursCounter_1.TcDUT
//   POUs/Tc3 Objects/Measurements/ FB_MeanValue.TcPOU, FB_TemperaturOK_1.TcPOU, FB_Timer_1.TcPOU, ST_Time_1.TcDUT
//   POUs/Tc3 Objects/Measurements/Oscat/ T_PLC_MS_1.TcPOU
//   POUs/Tc3 Objects/Measurements/RTC/ FB_RTC_1.TcPOU
//   POUs/Tc3 Objects/Safety/ FB_AirPressure_1.TcPOU, FB_LightCurtain_1.TcPOU, FB_NoEmergencyStop_1.TcPOU, FB_PowerSupply_1.TcPOU, FB_Temperature_1.TcPOU
//   POUs/Tc3 Objects/Safety/Fieldbus/EtherCAT Diag/ ET_EtherCATDiag_1.TcDUT (not stored), E_EcCommState_1.TcDUT (not stored), FB_EtherCATDiag_1.TcPOU (not stored), FB_EtherCATFrameDiag_1.TcPOU (not stored), ST_EcMasterDevState_1.TcDUT (not stored), ST_SlaveStateInfoScanned_1.TcDUT (not stored), ST_SlaveStateInfo_1.TcDUT (not stored), ST_SlaveState_1.TcDUT (not stored), ST_TopologyData_1.TcDUT (not stored)
//   POUs/Tc3 Objects/Safety/Fieldbus/ FB_Fieldbus_1.TcPOU, ST_FieldbusStatus_1.TcDUT
//   POUs/Tc3 Objects/Signals/Force Input/ FB_ForceBit_1.TcPOU, FB_ForceByte_1.TcPOU, FB_ForceInput.TcPOU
//   POUs/Tc3 Objects/Signals/Generators/ FB_Blinker_1.TcPOU, ST_Blinker_1.TcDUT
//   POUs/Tc3 Objects/Signals/Handling/ FB_SignalHandlingDelay_1.TcPOU, FB_SignalHandlingEdge_1.TcPOU, F_SignalHandling_1.TcPOU
//   POUs/Tc3 Objects/Signals/Ramp Generators/ ET_RampGenerator_1.TcDUT, FB_RampDirector_1.TcPOU
//   POUs/Tc3 Objects/Signals/Ramp Generators/Oscat_Ramp/ FB_RMP_W_1.TcPOU (not stored), _RMP_W_1.TcPOU (not stored)
//   POUs/Tc3 Objects/Signals/Watchdog/ FB_SignalWatchdogLimit.TcPOU, FB_SignalWatchdog_1.TcPOU
//   POUs/Tc3 Objects/String/ F_CheckStringIsReal_1.TcPOU, F_CheckSyntaxReal.TcPOU, F_CheckSyntaxString.TcPOU, F_RealToStrf_1.TcPOU
//   POUs/Tc3 Objects/Traceability/ ET_TRACE_State.TcDUT, FB_TraceCycle.TcPOU, FB_TraceSingle.TcPOU, GVL_Trace.TcGVL

CONFIGURATION _49001_01_BSM_762_V01_000_ISCOtherm
    RESOURCE PLC ON TwinCAT3
        TASK PLC_TASK(INTERVAL := T#10ms, PRIORITY := 1);
        PROGRAM MAIN WITH PLC_TASK : MAIN;
    END_RESOURCE
END_CONFIGURATION

// ---- Data types/Machine/BECKHOFF/ST_BECKHOFFDRIVETOPLC.TcDUT
(* Communication structure from drive to plc *)

TYPE ST_BECKHOFFDRIVETOPLC :
STRUCT
	bAxisHELimitMax 					:BOOL; 						(* DI1.7 Maximum limit of  axis heating element / Endschalter Achse Heizelement maximal *)
	bAxisHELimitMin 					:BOOL;						(* DI1.6 Minimum limit of  axis heating element / Endschalter Achse Heizelement minimal *)
END_STRUCT
END_TYPE

// ---- Data types/Machine/BECKHOFF/ST_BECKHOFFDRIVE_REF.TcDUT
TYPE ST_BECKHOFFDRIVE_REF : FB_BECKHOFFDRIVE_REF;
END_TYPE

// ---- Data types/Machine/BECKHOFF/ST_PLCTOBECKHOFFDRIVE.TcDUT
(* Communication structure from plc to drive *)

TYPE ST_PLCTOBECKHOFFDRIVE :
STRUCT
		wPO1ControlWord						:WORD;
END_STRUCT
END_TYPE

// ---- Data types/Machine/FORCE/ST_FORCETOPLC.TcDUT
(* Communication structure from drive to plc *)

TYPE ST_FORCETOPLC :
STRUCT

END_STRUCT
END_TYPE

// ---- Data types/Machine/FORCE/ST_FORCE_REF.TcDUT
TYPE ST_FORCE_REF : FB_FORCE_REF;
END_TYPE

// ---- Data types/Machine/FORCE/ST_PLCTOFORCE.TcDUT
(* Communication structure from plc to drive *)

TYPE ST_PLCTOFORCE :
STRUCT

END_STRUCT
END_TYPE

// ---- Data types/Machine/Group_0000 - General/ET_Gr00Auto.TcDUT
TYPE ET_Gr00Auto :
(
	ET_Gr00Auto_eWaitExecute := 0,
	ET_Gr00Auto_eAutomatic,
	ET_Gr00Auto_eInterrupted := 196,
	ET_Gr00Auto_eDone := 197,
	ET_Gr00Auto_eError := 198,
	ET_Gr00Auto_eNoExecute := 199
);
END_TYPE

// ---- Data types/Machine/Group_0000 - General/ET_Gr00Home.TcDUT
TYPE ET_Gr00Home :
(
	ET_Gr00Home_eWaitExecute := 0,
	ET_Gr00Home_eReference,
	ET_Gr00Home_eReadPrg,
	ET_Gr00Home_eWfReadPrg,
	ET_Gr00Home_eProgramVerification,
	ET_Gr00Home_eWfErrorByProgramVerification,
	ET_Gr00Home_eDone := 197,
	ET_Gr00Home_eError := 198,
	ET_Gr00Home_eNoExecute := 199
);
END_TYPE

// ---- Data types/Machine/Group_0000 - General/ST_Gr00HMIRef.TcDUT
TYPE ST_Gr00HMIRef :
STRUCT
	stHMITOPLC				:ST_Gr00HMITOPLC;
	stPLCTOHMI				:ST_Gr00PLCTOHMI;
END_STRUCT
END_TYPE

// ---- Data types/Machine/Group_0000 - General/ST_Gr00HMITOPLC.TcDUT
TYPE ST_Gr00HMITOPLC :
STRUCT
	etMachineMode			:ET_MachineMode;			(* Machine mode enum variable *)
	bBtnStart					:BOOL; 						(* Button start *)
	bBtnStop					:BOOL; 						(* Button stop *)
	bBtnReset				:BOOL; 						(* Button reset *)
	bBtnForceRef				:BOOL; 						(* Button reference force *)
	bBtnMachinePurge		:BOOL;						(* Button machine purge  *)
	bResetCounterUser		:BOOL;						(* Reset counter user *)
	bSafetyInterlockOff		:BOOL;						(* Deactivation safety interlocks if machine is in manual mode *)
	bProgramActive			:BOOL;						(* Program active *)
	rOverride				:REAL;						(* Override *)
	sActRecipe 				:STRING;					(* Current recipe *)
END_STRUCT
END_TYPE

// ---- Data types/Machine/Group_0000 - General/ST_Gr00PLCTOHMI.TcDUT
TYPE ST_Gr00PLCTOHMI :
STRUCT
	etMachineMode						:ET_MachineMode;			(* Machine mode *)
	etMachineState						:ET_MachineState;			(* Machine state *)
	wBtnStartStatus						:WORD;						(* Button start status *)
	wBtnStopStatus						:WORD;						(* Button stop status *)
	wBtnResetStatus						:WORD;						(* Button reset status *)
	wBtnForceRefStatus					:WORD;						(* Button reference force status *)
	wBtnAutoStatus						:WORD;						(* Button auto status *)
	wBtnHomeStatus						:WORD;						(* Button home status *)
	wBtnManualStatus						:WORD;						(* Button manual status *)
	wLampStatus							:WORD;						(* Lamp status *)
	wAlarmStatus							:WORD;						(* Alarm status *)
	bMachineRunning						:BOOL;						(* Machine running *)
	bHomeCompleted						:BOOL;						(* Home completed *)
	bAutoCompleted						:BOOL;						(* Auto completed *)
	bModeAutomatic						:BOOL;						(* Machine mode automatic *)
	bModeHome							:BOOL;						(* Machine mode home *)
	bModeManual						:BOOL;						(* Machine mode manual *)
	udnCounterTotal						:UDINT;						(* Total counter *)
	udnCounterUser						:UDINT;						(* User counter *)
	dwCycleTime							:DWORD;					(* Cycletime in 0.01sec / Zykluszeit in 0.01Sekunden *)
	lrMachineLifetime						:LREAL;				 		(* Machine lifetime *)
	lrMachineLifetimeAfterTurnOn			:LREAL;				 		(* Machine lifetime after turn on *)
	sPrgFilePath							:STRING;					(* Current program file path *)
END_STRUCT
END_TYPE

// ---- Data types/Machine/Group_0001/ET_Gr01Auto.TcDUT
TYPE ET_Gr01Auto :
(
	ET_Gr01Auto_eWaitExecute := 0,
	ET_Gr01Auto_eWaitAxisStatus,
	ET_Gr01Auto_eGetProcessPara,
	ET_Gr01Auto_eWfErrorCollisionDetected,
	ET_Gr01Auto_eChkProcessEnd,
	ET_Gr01Auto_eAxisAngleToWorkPos,
	ET_Gr01Auto_eWfAxisAngleInWorkPos,
	ET_Gr01Auto_eWfReq,
	ET_Gr01Auto_eAngleAck,
	ET_Gr01Auto_eSawingAck,
	ET_Gr01Auto_eSawbandStart,
	ET_Gr01Auto_eWfSawbandStart,
	ET_Gr01Auto_eSawingStart,
	ET_Gr01Auto_eWfSawingDone,
	ET_Gr01Auto_eAxisSawBowToSafePos,
	ET_Gr01Auto_eWfAxisSawBowInSafePos,
	ET_Gr01Auto_eStopOrContinue,
	ET_Gr01Auto_eSawBandStop,
	ET_Gr01Auto_eSawBandStopped,
	ET_Gr01Auto_eTransportReq,
	ET_Gr01Auto_eTransportAck,
	ET_Gr01Auto_eAxisSawBowToSafePos2,
	ET_Gr01Auto_eWfAxisSawBowInSafePos2,
	ET_Gr01Auto_eAxisAngleToBasePos,
	ET_Gr01Auto_eWfAxisAngleInBasePos,
	ET_Gr01Auto_eDone := 197,
	ET_Gr01Auto_eError := 198,
	ET_Gr01Auto_eNoExecute := 199
);
END_TYPE

// ---- Data types/Machine/Group_0001/ET_Gr01Home.TcDUT
TYPE ET_Gr01Home :
(
	ET_Gr01Home_eWaitExecute := 0,
	ET_Gr01Home_eWaitAxisStatus,
	ET_Gr01Home_eGetProcessPara,
	ET_Gr01Home_eSawbandStop,
	ET_Gr01Home_eWfSawbandStopped,
	ET_Gr01Home_eAxisSawbandGuide,
	ET_Gr01Home_eWfAxisSawbandGuide,
	ET_Gr01Home_eAxisSawBow,
	ET_Gr01Home_eWfAxisSawBow,
	ET_Gr01Home_eAxisAngle,
	ET_Gr01Home_eWfAxisAngle,
	ET_Gr01Home_eWfFreeToMove,
	ET_Gr01Home_eAxisSawBowMoveHomePos,
	ET_Gr01Home_eWfAxisSawBowInHomePos,
	ET_Gr01Home_eDone := 197,
	ET_Gr01Home_eError := 198,
	ET_Gr01Home_eNoExecute := 199
);
END_TYPE

// ---- Data types/Machine/Group_0001/ET_Gr01HomeAxis.TcDUT
TYPE ET_Gr01HomeAxis :
(
	ET_Gr01HomeAxis_eWaitExecute := 0,
	ET_Gr01HomeAxis_eWaitAxisStatus,
	ET_Gr01HomeAxis_eMoveStop,
	ET_Gr01HomeAxis_eWFMoveStop,
	ET_Gr01HomeAxis_eAxisReset,
	ET_Gr01HomeAxis_eWfAxisReset,
	ET_Gr01HomeAxis_eChkAxisCoupled,
	ET_Gr01HomeAxis_eAxisRef,
	ET_Gr01HomeAxis_eWfAxisRef,
	ET_Gr01HomeAxis_eWfErrorByReference,
	ET_Gr01HomeAxis_eAxisMoveHomePos,
	ET_Gr01HomeAxis_eAxisInHomePos,
	ET_Gr01HomeAxis_eAxisSetHome,
	ET_Gr01HomeAxis_eWfSetHome,
	ET_Gr01HomeAxis_eDone := 197,
	ET_Gr01HomeAxis_eError := 198,
	ET_Gr01HomeAxis_eNoExecute := 199
);
END_TYPE

// ---- Data types/Machine/Group_0001/ET_Gr01HomeSawband.TcDUT
TYPE ET_Gr01HomeSawband :
(
	ET_Gr01HomeSawband_eWaitExecute := 0,
	ET_Gr01HomeSawband_eStop,
	ET_Gr01HomeSawband_eWFStop,
	ET_Gr01HomeSawband_eReset,
	ET_Gr01HomeSawband_eWfReset,
	ET_Gr01HomeSawband_eDone := 197,
	ET_Gr01HomeSawband_eError := 198,
	ET_Gr01HomeSawband_eNoExecute := 199
);
END_TYPE

// ---- Data types/Machine/Group_0001/ET_Gr01Manual.TcDUT
TYPE ET_Gr01Manual :
(
	ET_Gr01Manual_eWaitExecute := 0,
	ET_Gr01Manual_eSetPosAxis5,
	ET_Gr01Manual_eWfSetPosAxis5,
	ET_Gr01Manual_eCouplingAxis1_4,
	ET_Gr01Manual_eWfCouplingAxis1_4,
	ET_Gr01Manual_eDone := 197,
	ET_Gr01Manual_eError := 198,
	ET_Gr01Manual_eNoExecute := 199
);
END_TYPE

// ---- Data types/Machine/Group_0001/ST_Gr01HMIRef.TcDUT
TYPE ST_Gr01HMIRef :
STRUCT
	stHMITOPLC				:ST_Gr01HMITOPLC;
	stPLCTOHMI				:ST_Gr01PLCTOHMI;
END_STRUCT
END_TYPE

// ---- Data types/Machine/Group_0001/ST_Gr01HMITOPLC.TcDUT
TYPE ST_Gr01HMITOPLC :
STRUCT
	bBtnStart							:BOOL; 											(* Button start *)
	bBtnStop							:BOOL; 											(* Button stop *)
	bBtnSteppingProcess					:BOOL; 											(* Stepping process *)
	rOverride							:REAL;											(* Override 0 - 100 [%]  *)
	bResetLifetime						:BOOL;											(* Reset life time *)
   	bResetCounterUser				   	:BOOL;											(* Reset counter user *)
	bBtnAxisSawBowPlus					:BOOL;											(* Button move axis saw bow plus *)
	bBtnAxisSawBowMinus					:BOOL;											(* Button move axis saw bow minus *)
	bBtnAxisAnglePlus					:BOOL;											(* Button move axis angle plus *)
	bBtnAxisAngleMinus					:BOOL;											(* Button move axis angle minus *)
	bBtnSawbandPlus						:BOOL;											(* Button saw band plus *)
	bBtnSawbandMinus					:BOOL;											(* Button saw band minus *)
	bBtnSawbandAirOn					:BOOL;											(* On sawband air *)
	bBtnSawbandAirOff					:BOOL;											(* Off sawband air *)
	bBtnLaserOn							:BOOL;											(* On laser *)
	bBtnLaserOff						:BOOL;											(* Off laser *)
	bBtnVacuumCleanerOn					:BOOL;											(* Vacuum cleaner on *)
	bBtnVacuumCleanerOff				:BOOL;											(* Vacuum cleaner off *)
	lrAxisSawBowTipDistance				:LREAL;											(* Tip distance axis saw bow [mm] *)
	lrAxisSawBowOriginShiftPos			:LREAL;											(* Origin shift position axis saw bow [mm] *)
	lrAxisSawBowHomePos					:LREAL;											(* Home position axis saw bow [mm] *)
	lrAxisSawBowSoftLimitMax			:LREAL;											(* Software limit maximum axis saw bow [mm] *)
	lrAxisSawBowSoftLimitMin			:LREAL;											(* Software limit minimum axis saw bow [mm] *)
	lrAxisSawBowNoRefVelo				:LREAL;											(* No reference velocity axis saw bow [%] *)
	lrAxisSawBowManualVelo				:LREAL;											(* Manual velocity axis saw bow [%] *)
	lrAxisSawBowHomeVelo				:LREAL;											(* Home velocity axis saw bow [%] *)
	lrAxisSawBowAutoVelo				:LREAL;											(* Auto velocity axis saw bow [%] *)
	lrAxisAngleTipDistance				:LREAL;											(* Tip distance axis angle [mm] *)
	lrAxisAngleOriginShiftPos			:LREAL;											(* Origin shift position axis angle [mm] *)
	lrAxisAngleHomePos					:LREAL;											(* Home position axis angle [mm] *)
	lrAxisAngleSoftLimitMax				:LREAL;											(* Software limit maximum axis angle [mm] *)
	lrAxisAngleSoftLimitMin				:LREAL;											(* Software limit minimum axis angle [mm] *)
	lrAxisAngleNoRefVelo				:LREAL;											(* No reference velocity axis angle [%] *)
	lrAxisAngleManualVelo				:LREAL;											(* Manual velocity axis angle [%] *)
	lrAxisAngleHomeVelo					:LREAL;											(* Home velocity axis angle [%] *)
	lrAxisAngleAutoVelo					:LREAL;											(* Auto velocity axis angle [%] *)
	rSawbandManualSpeed					:REAL;											(* Manual speed sawband [upm] *)
	rSawbandAutoSpeed					:REAL;											(* Auto speed sawband [upm] *)
	rSawingOverride						:REAL;											(* Sawing override 0 - 100 [%]  *)
	rPipeDiameter						:REAL;											(* Pipe diameter [mm] *)
	lrActSawingAngle					:LREAL;											(* Actual angle of sawing [mm] *)
	lrSafetyDistance					:LREAL;											(* Safety distance [mm] *)
	lrSafeDistSawBandToPipe				:LREAL;											(* Safety distance sawband to pipe[mm] *)
	lrSawBandThickness					:LREAL;											(* Sawband thickness [mm] *)
END_STRUCT
END_TYPE

// ---- Data types/Machine/Group_0001/ST_Gr01PLCTOHMI.TcDUT
TYPE ST_Gr01PLCTOHMI :
STRUCT
	wBtnStartStatus						:WORD;						(* Button start status *)
	wBtnStopStatus						:WORD;						(* Button stop status *)
	wBtnStepProcStatus					:WORD;						(* Button stepping process status *)
	bHomeCompleted						:BOOL;						(* Home completed *)
	bExecutedProcess					:BOOL;						(* Process executed *)
	udnCounterTotal						:UDINT;						(* Total counter *)
	dwCycleTime							:DWORD;					(* Cycletime in 0.01sec / Zykluszeit in 0.01Sekunden *)
	lrLifetime							:LREAL;				 		(* Lifetime *)
	lrLifetimeAfterReset				:LREAL;				 		(* Lifetime after reset *)
	lrLifetimeAfterTurnOn				:LREAL;				 		(* Lifetime after turn on *)
	wAxisSawBowStatus					:WORD;						(* Axis saw bow status *)
	wAxisAngleStatus					:WORD;						(* Axis angle status *)
	wSawbandStatus						:WORD;						(* Sawband status *)
    wSawbandAirStatus 					:WORD;						(* Sawband air status *)
    wLaserStatus						:WORD;                 				(* Sawband laser status *)
	lrAxisSawBowActPos					:LREAL;						(* Axis saw bow actual position *)
	lrAxisSawBowActVelo					:LREAL;						(* Axis saw bow actual velocity *)
	lrAxisSawBowActForce				:LREAL;						(* Axis saw bow actual force *)
	lrAxisAngleActPos					:LREAL;						(* Axis angle actual position *)
	lrAxisAngleActVelo					:LREAL;						(* Axis angle actual velocity *)
	lrAxisAngleActForce					:LREAL;						(* Axis angle actual force *)
	lrSawbandActSpeed					:LREAL;						(* Actual speed of sawband *)
END_STRUCT
END_TYPE

// ---- Data types/Machine/Group_0002/ET_Gr02Auto.TcDUT
TYPE ET_Gr02Auto :
(
	ET_Gr02Auto_eWaitExecute := 0,
	ET_Gr02Auto_eWaitAxisStatus,
	ET_Gr02Auto_eGetPart,
	ET_Gr02Auto_eFixPart,
	ET_Gr02Auto_eWarrningPartNoPresent,
	ET_Gr02Auto_eStartProgramReq,
	ET_Gr02Auto_eStartProgramAck,
	ET_Gr02Auto_eAxisRef,
	ET_Gr02Auto_eWfAxisRef,
	ET_Gr02Auto_eDelayStartSection,
	ET_Gr02Auto_eWfDelayStartSection,
	ET_Gr02Auto_eStartSection,
	ET_Gr02Auto_eStopExtruderReq,
	ET_Gr02Auto_eWfStartSection,
	ET_Gr02Auto_eReleasePart,
	ET_Gr02Auto_eDone := 197,
	ET_Gr02Auto_eError := 198,
	ET_Gr02Auto_eNoExecute := 199
);
END_TYPE

// ---- Data types/Machine/Group_0002/ET_Gr02Home.TcDUT
TYPE ET_Gr02Home :
(
	ET_Gr02Home_eWaitExecute := 0,
	ET_Gr02Home_eWaitAxisStatus,
	ET_Gr02Home_eHomePreparation,
	ET_Gr02Home_eChkHomeMode,
	ET_Gr02Home_eWfFreeToMove,
	ET_Gr02Home_eCylinderToBase,
	ET_Gr02Home_eAxisClamping,
	ET_Gr02Home_eWfAxisClamping,
	ET_Gr02Home_eDone := 197,
	ET_Gr02Home_eError := 198,
	ET_Gr02Home_eNoExecute := 199
);
END_TYPE

// ---- Data types/Machine/Group_0002/ET_Gr02HomeAxis.TcDUT
TYPE ET_Gr02HomeAxis :
(
	ET_Gr02HomeAxis_eWaitExecute := 0,
	ET_Gr02HomeAxis_eWaitAxisStatus,
	ET_Gr02HomeAxis_eMoveStop,
	ET_Gr02HomeAxis_eWFMoveStop,
	ET_Gr02HomeAxis_eAxisReset,
	ET_Gr02HomeAxis_eWfAxisReset,
	ET_Gr02HomeAxis_eChkAxisCoupled,
	ET_Gr02HomeAxis_eAxisRef,
	ET_Gr02HomeAxis_eWfAxisRef,
	ET_Gr02HomeAxis_eWfErrorByReference,
	ET_Gr02HomeAxis_eAxisMoveHomePos,
	ET_Gr02HomeAxis_eAxisInHomePos,
	ET_Gr02HomeAxis_eAxisSetHome,
	ET_Gr02HomeAxis_eWfSetHome,
	ET_Gr02HomeAxis_eDone := 197,
	ET_Gr02HomeAxis_eError := 198,
	ET_Gr02HomeAxis_eNoExecute := 199
);
END_TYPE

// ---- Data types/Machine/Group_0002/ET_Gr02Manual.TcDUT
TYPE ET_Gr02Manual :
(
	ET_Gr02Manual_eWaitExecute := 0,
	ET_Gr02Manual_eSetPosAxis5,
	ET_Gr02Manual_eWfSetPosAxis5,
	ET_Gr02Manual_eCouplingAxis1_4,
	ET_Gr02Manual_eWfCouplingAxis1_4,
	ET_Gr02Manual_eDone := 197,
	ET_Gr02Manual_eError := 198,
	ET_Gr02Manual_eNoExecute := 199
);
END_TYPE

// ---- Data types/Machine/Group_0002/ST_Gr02HMIRef.TcDUT
TYPE ST_Gr02HMIRef :
STRUCT
	stHMITOPLC				:ST_Gr02HMITOPLC;
	stPLCTOHMI				:ST_Gr02PLCTOHMI;
END_STRUCT
END_TYPE

// ---- Data types/Machine/Group_0002/ST_Gr02HMITOPLC.TcDUT
TYPE ST_Gr02HMITOPLC :
STRUCT
	bBtnStart								:BOOL; 											(* Button start *)
	bBtnStop								:BOOL; 											(* Button stop *)
	bBtnSteppingProcess					:BOOL; 											(* Stepping process *)
	rOverride							:REAL;											(* Override 0 - 100 [%]  *)
	bResetLifetime						:BOOL;											(* Reset life time *)
         bResetCounterUser			   		:BOOL;											(* Reset counter user *)
END_STRUCT
END_TYPE

// ---- Data types/Machine/Group_0002/ST_Gr02PLCTOHMI.TcDUT
TYPE ST_Gr02PLCTOHMI :
STRUCT
	wBtnStartStatus						:WORD;						(* Button start status *)
	wBtnStopStatus						:WORD;						(* Button stop status *)
	wBtnStepProcStatus					:WORD;						(* Button stepping process status *)
	bHomeCompleted						:BOOL;						(* Home completed *)
	bExecutedProcess					:BOOL;						(* Process executed *)
	udnCounterTotal						:UDINT;						(* Total counter *)
	dwCycleTime							:DWORD;					(* Cycletime in 0.01sec / Zykluszeit in 0.01Sekunden *)
	lrLifetime								:LREAL;				 		(* Lifetime *)
	lrLifetimeAfterReset					:LREAL;				 		(* Lifetime after reset *)
	lrLifetimeAfterTurnOn					:LREAL;				 		(* Lifetime after turn on *)
END_STRUCT
END_TYPE

// ---- Data types/Machine/Group_0005/ET_Gr05Auto.TcDUT
TYPE ET_Gr05Auto :
(
	ET_Gr05Auto_eWaitExecute := 0,
	ET_Gr05Auto_eWaitAxisStatus,
	ET_Gr05Auto_eClamp1Close,
	ET_Gr05Auto_ChkPipeBeginEdge,
	ET_Gr05Auto_eAxisClamp1InPipeBeginPos,
	ET_Gr05Auto_eClamp2Open,
	ET_Gr05Auto_eAxisClamp1MoveVeloPipeBegin,
	ET_Gr05Auto_eWfAxisClamp1MoveVeloPipeBegin,
	(*ET_Gr05Auto_eAxisClamp1InPipeBeginPos,*)
	ET_Gr05Auto_eGetClamp1ActPos,
	ET_Gr05Auto_eWfPipeBeginNoDetectedError,
	ET_Gr05Auto_eWfPipeBeginNoDetectedWarrning,
	ET_Gr05Auto_eEnd,
	ET_Gr05Auto_eSawbandStart,
	ET_Gr05Auto_eAxisClamp1MoveToSawBandPos,
	ET_Gr05Auto_eAxisClamp1InSawBandPos,
	ET_Gr05Auto_eAxisClamp2MoveToSawBandPos,
	ET_Gr05Auto_eAxisClamp2InSawBandPos,
	ET_Gr05Auto_eGetClamp1ActPos_01,
	ET_Dummy_01A,
	ET_Dummy_01B,
	ET_Gr05Auto_eAxisClamp2MoveSawPos,
	ET_Gr05Auto_eAxisClamp2InSawPos,
	ET_Gr05Auto_eGetProcessPara,
	ET_Gr05Auto_eChkProcessEnd,
	ET_Gr05Auto_eClamp12Open,
	(*ET_Gr05Auto_eEnd,*)
	ET_Gr05Auto_eWfSlideUp,
	ET_Gr05Auto_eGetClamp2ActPos,
	ET_Gr05Auto_eCollisionDetectedErr,
	ET_Gr05Auto_eChkWorkArea,

	ET_Gr05Auto_ChkPipeEndDetected,
	(*ET_Gr05Auto_eClamp12Open,*)
	ET_Gr05Auto_eClamp2Close,
	ET_Gr05Auto_eClamp2CloseErr,
	ET_Gr05Auto_eClamp1Open,
	ET_Gr05Auto_eClamp1OpenErr,
	ET_Gr05Auto_eAxisClamp1MoveAbsPipeEnde,
	ET_Gr05Auto_eAxisClamp1MoveAbsPipeEndeErr,

	ET_Gr05Auto_eWfAxisClamp1MoveAbsPipeEnde,(*pipe end detected*)

	ET_Gr05Auto_eGetClamp1ActPos_03,
	ET_Gr05Auto_eClamp1Close3,
	ET_Gr05Auto_eChkAdjustSawingLength,
	(*ET_Gr05Auto_eChkProcessEnd,*)
	ET_Gr05Auto_NurWennlrActRemoveLength_0,
	ET_Gr05Auto_eClamp2Open3,
	ET_Gr05Auto_eAxisClamp2MoveToPos2,
	ET_Gr05Auto_eAxisClamp2InPos2,
	ET_Gr05Auto_eAxisClamp1MoveToPos2,
	ET_Gr05Auto_eAxisClamp1InPos2,
	ET_Gr05Auto_eSawingLengthCorrection,
	(*ET_Gr05Auto_ChkPipeEndDetected,*)


	ET_Gr05Auto_eAxisClamp1Stop,
	ET_Gr05Auto_eWfAxisClamp1Stop,
	ET_Gr05Auto_eGetClamp1ActPos_04,
	ET_Gr05Auto_eChkNextSawingAngle,

	ET_Gr05Auto_eAxisClamp1MoveVeloPipeEnd,
	ET_Gr05Auto_eWfAxisClamp1MoveVeloPipeEnd,
	ET_Gr05Auto_eAxisClamp1InPipeEndPos,
	ET_Gr05Auto_eWfPipeEndNoDetectedErr,
	ET_Gr05Auto_eAxisClamp1Stop_2,
	ET_Gr05Auto_eAxisClamp1StopErr_2,
	ET_Gr05Auto_eWfAxisClamp1Stop_2,
	ET_Gr05Auto_eWfAxisClamp1StopErr_2,

	ET_Gr05Auto_ChkNextSawingLenght,
	ET_Gr05Auto_eGetClamp1ActPos_05,
	ET_Gr05Auto_eAngleReq,
	ET_Gr05Auto_eAngleAck,
	Dummy_03,
	(*ET_Gr05Auto_eChkProcessEnd,*)


	ET_Gr05Auto_eAxisClamp1StopErr,

	(*ET_Gr05Auto_eGetClamp1ActPos_03,*)
	ET_Gr05Auto_eWfAxisClamp1MoveAbsPipeEndeErr,



	ET_Gr05Auto_eClamp1Close2,
	ET_Gr05Auto_eClamp2Open1,
	ET_Gr05Auto_eAxisClamp1MoveToPos,
	ET_Gr05Auto_eAxisClamp1InPos,
	ET_Gr05Auto_eAxisClamp2MoveToPos,
	ET_Gr05Auto_eAxisClamp2InPos,
	ET_Gr05Auto_eGetClamp1ActPos_02,
	ET_Dummy_02A,
	ET_Dummy_02B,
	ET_Gr05Auto_eChkAxisClamp1MoveToBackPos,
	ET_Gr05Auto_eClamp2Slide,
	ET_Gr05Auto_eClamp2Err,
	ET_Gr05Auto_eSlideUpErr,

	ET_Gr05Auto_eAxisClamp1MoveToBackPos,
	ET_Gr05Auto_eAxisClamp1MoveToBackPosErr,
	ET_Gr05Auto_eAxisClamp1InBackPos,
	ET_Gr05Auto_eGetClamp1ActPos_06,
	(*ET_Gr05Auto_eChkProcessEnd,*)
	ET_Gr05Auto_eAxisClamp1InBackPosErr,


	ET_Gr05Auto_eSawingReq,
	ET_Gr05Auto_eSawingAck,
	ET_Gr05Auto_eWfTransportReq,
	ET_Gr05Auto_eTransportAck,
	ET_Gr05Auto_eSlideDown,
	ET_Gr05Auto_eSlideDownErr,
	ET_Gr05Auto_eRemovalBandErr,

	ET_Gr05Auto_eInterrupted := 196,
	ET_Gr05Auto_eDone := 197,
	ET_Gr05Auto_eError := 198,
	ET_Gr05Auto_eNoExecute := 199
);
END_TYPE

// ---- Data types/Machine/Group_0005/ET_Gr05AutoProcess.TcDUT
TYPE ET_Gr05AutoProcess :
(
	ET_Gr05AutoProcess_eWaitExecute := 0,
	ET_Gr05AutoProcess_eWaitAxisStatus,
	ET_Gr05AutoProcess_eWfStartProcessReq,
	ET_Gr05AutoProcess_eStartProcessPrg,
	ET_Gr05AutoProcess_eWfProcessPrgDone,
	ET_Gr05AutoProcess_eExtruderStart,
	ET_Gr05AutoProcess_eWfExtruderStart,
	ET_Gr05AutoProcess_eExtruderStop,
	ET_Gr05AutoProcess_eWfExtruderStop,
	ET_Gr05AutoProcess_eStartEndPrg,
	ET_Gr05AutoProcess_eWfEndPrgDone,
	ET_Gr05AutoProcess_ePrgInterrupted,
	ET_Gr05AutoProcess_eStartHomePrg,
	ET_Gr05AutoProcess_eWfHomePrgDone,
	ET_Gr05AutoProcess_eInterrupted := 196,
	ET_Gr05AutoProcess_eDone := 197,
	ET_Gr05AutoProcess_eError := 198,
	ET_Gr05AutoProcess_eNoExecute := 199
);
END_TYPE

// ---- Data types/Machine/Group_0005/ET_Gr05Home.TcDUT
TYPE ET_Gr05Home :
(
	ET_Gr05Home_eWaitExecute := 0,
	ET_Gr05Home_eWaitAxisStatus,
	ET_Gr05Home_eWfFreeToMove,
	ET_Gr05Home_eClampsSlide,
	ET_Gr05Home_eAxisClamp1,
	ET_Gr05Home_eWfAxisClamp1,
	ET_Gr05Home_eAxisClamp2,
	ET_Gr05Home_eWfAxisClamp2,
	ET_Gr05Home_eDone := 197,
	ET_Gr05Home_eError := 198,
	ET_Gr05Home_eNoExecute := 199
);
END_TYPE

// ---- Data types/Machine/Group_0005/ET_Gr05HomeAxis.TcDUT
TYPE ET_Gr05HomeAxis :
(
	ET_Gr05HomeAxis_eWaitExecute := 0,
	ET_Gr05HomeAxis_eWaitAxisStatus,
	ET_Gr05HomeAxis_eMoveStop,
	ET_Gr05HomeAxis_eWFMoveStop,
	ET_Gr05HomeAxis_eAxisReset,
	ET_Gr05HomeAxis_eWfAxisReset,
	ET_Gr05HomeAxis_eChkAxisCoupled,
	ET_Gr05HomeAxis_eAxisRef,
	ET_Gr05HomeAxis_eWfAxisRef,
	ET_Gr05HomeAxis_eWfErrorByReference,
	ET_Gr05HomeAxis_eAxisMoveHomePos,
	ET_Gr05HomeAxis_eAxisInHomePos,
	ET_Gr05HomeAxis_eAxisSetHome,
	ET_Gr05HomeAxis_eWfSetHome,
	ET_Gr05HomeAxis_eDone := 197,
	ET_Gr05HomeAxis_eError := 198,
	ET_Gr05HomeAxis_eNoExecute := 199
);
END_TYPE

// ---- Data types/Machine/Group_0005/ET_Gr05HomeAxisClamp1.TcDUT
TYPE ET_Gr05HomeAxisClamp1 :
(
	ET_Gr05HomeAxisClamp1_eWaitExecute := 0,
	ET_Gr05HomeAxisClamp1_eWaitAxisStatus,
	ET_Gr05HomeAxisClamp1_eMoveStop,
	ET_Gr05HomeAxisClamp1_eWFMoveStop,
	ET_Gr05HomeAxisClamp1_eAxisReset,
	ET_Gr05HomeAxisClamp1_eWfAxisReset,
	ET_Gr05HomeAxisClamp1_eChkAxisCoupled,
	ET_Gr05HomeAxisClamp1_eAxisRef,
	ET_Gr05HomeAxisClamp1_eWfAxisRef,
	ET_Gr05HomeAxisClamp1_eWfErrorByReference,
	ET_Gr05HomeAxisClamp1_eWfErrorByPipeCollision,
	ET_Gr05HomeAxisClamp1_eAxisMoveHomePos,
	ET_Gr05HomeAxisClamp1_eAxisInHomePos,
	ET_Gr05HomeAxisClamp1_eMoveStop2,
	ET_Gr05HomeAxisClamp1_eWFMoveStop2,
	ET_Gr05HomeAxisClamp1_eAxisMovePipeEndVelo,
	ET_Gr05HomeAxisClamp1_eWfAxisInPipeEndVelo,
	ET_Gr05HomeAxisClamp1_eMoveStop3,
	ET_Gr05HomeAxisClamp1_eWFMoveStop3,
	ET_Gr05HomeAxisClamp1_eWfErrorByPipeEndNoDetected,
	ET_Gr05HomeAxisClamp1_eDone := 197,
	ET_Gr05HomeAxisClamp1_eError := 198,
	ET_Gr05HomeAxisClamp1_eNoExecute := 199
);
END_TYPE

// ---- Data types/Machine/Group_0005/ET_Gr05Manual.TcDUT
TYPE ET_Gr05Manual :
(
	ET_Gr05Manual_eWaitExecute := 0,
	ET_Gr05Manual_eDone := 197,
	ET_Gr05Manual_eError := 198,
	ET_Gr05Manual_eNoExecute := 199
);
END_TYPE

// ---- Data types/Machine/Group_0005/ST_Gr05HMIRef.TcDUT
TYPE ST_Gr05HMIRef :
STRUCT
	stHMITOPLC				:ST_Gr05HMITOPLC;
	stPLCTOHMI				:ST_Gr05PLCTOHMI;
END_STRUCT
END_TYPE

// ---- Data types/Machine/Group_0005/ST_Gr05HMITOPLC.TcDUT
TYPE ST_Gr05HMITOPLC :
STRUCT
	bBtnStart								:BOOL; 											(* Button start *)
	bBtnStop								:BOOL; 											(* Button stop *)
	bBtnSteppingProcess					:BOOL; 											(* Stepping process *)
	rOverride							:REAL;											(* Override 0 - 100 [%]  *)
	bResetLifetime						:BOOL;											(* Reset life time *)
         bResetCounterUser			   		:BOOL;											(* Reset counter user *)
	arbBtnAxisClampPlus					:ARRAY[1..ungGr05ClampMaxNo] OF BOOL;			(* Button move axis clamp plus *)
	arbBtnAxisClampMinus					:ARRAY[1..ungGr05ClampMaxNo] OF BOOL;			(* Button move axis clamp minus *)
	arbBtnClampOpen						:ARRAY[1..ungGr05ClampMaxNo] OF BOOL;			(* Clamp open *)
	arbBtnClampClose					:ARRAY[1..ungGr05ClampMaxNo] OF BOOL;			(* Clamp close *)
	arbBtnCylinderPosOpen				:ARRAY[1..ungGr05CylinderPosMaxNo] OF BOOL;		(* Position cylinder open *)
	arbBtnCylinderPosClose				:ARRAY[1..ungGr05CylinderPosMaxNo] OF BOOL;		(* Position cylinder close *)
	bBtnSlideUp							:BOOL;											(* Button slide up *)
	bBtnSlideDown						:BOOL;											(* Button slide down *)
	bBtnRemovalBandToPlus				:BOOL;											(* Button move removal band into plus direction *)
	bBtnRemovalBandToMinus				:BOOL;											(* Button move removal band into minus direction *)
	bSlideActive							:BOOL;											(* Slide active *)
	bCylinderPosActive					:BOOL;											(* Position cylinder active *)
	arlrAxisClampTipDistance				:ARRAY[1..ungGr05ClampMaxNo] OF LREAL;			(* Tip distance axis clamp [mm] *)
	arlrAxisClampOriginShiftPos				:ARRAY[1..ungGr05ClampMaxNo] OF LREAL;			(* Origin shift position axis clamp [mm] *)
	arlrAxisClampHomePos				:ARRAY[1..ungGr05ClampMaxNo] OF LREAL;			(* Home position axis clamp [mm] *)
	arlrAxisClampSoftLimitMax				:ARRAY[1..ungGr05ClampMaxNo] OF LREAL;			(* Software limit maximum axis clamp [mm] *)
	arlrAxisClampSoftLimitMin				:ARRAY[1..ungGr05ClampMaxNo] OF LREAL;			(* Software limit minimum axis clamp [mm] *)
	arlrAxisClampNoRefVelo				:ARRAY[1..ungGr05ClampMaxNo] OF LREAL;			(* No reference velocity axis clamp [%] *)
	arlrAxisClampManualVelo				:ARRAY[1..ungGr05ClampMaxNo] OF LREAL;			(* Manual velocity axis clamp [%] *)
	arlrAxisClampHomeVelo				:ARRAY[1..ungGr05ClampMaxNo] OF LREAL;			(* Home velocity axis clamp [%] *)
	arlrAxisClampAutoVelo					:ARRAY[1..ungGr05ClampMaxNo] OF LREAL;			(* Auto velocity axis clamp [%] *)
	lrActSawingLength						:LREAL;											(* Actual sawing length [mm] *)
END_STRUCT
END_TYPE

// ---- Data types/Machine/Group_0005/ST_Gr05PLCTOHMI.TcDUT
TYPE ST_Gr05PLCTOHMI :
STRUCT
	wBtnStartStatus						:WORD;						(* Button start status *)
	wBtnStopStatus						:WORD;						(* Button stop status *)
	wBtnStepProcStatus					:WORD;						(* Button stepping process status *)
	bHomeCompleted						:BOOL;						(* Home completed *)
	bExecutedProcess					:BOOL;						(* Process executed *)
	udnCounterTotal						:UDINT;						(* Total counter *)
	dwCycleTime							:DWORD;					(* Cycletime in 0.01sec / Zykluszeit in 0.01Sekunden *)
	lrLifetime								:LREAL;				 		(* Lifetime *)
	lrLifetimeAfterReset					:LREAL;				 		(* Lifetime after reset *)
	lrLifetimeAfterTurnOn					:LREAL;				 		(* Lifetime after turn on *)
	wAxisClampStatus						:WORD;						(* Axis clamp 1 status *)
	wSlideStatus							:WORD;						(* Slide status *)
	wRemovalBandStatus					:WORD;						(* Removal band status *)
	arwClampStatus						:ARRAY[1..ungGr05ClampMaxNo] OF WORD;						(* Clamp status *)
	arwCylinderPosStatus					:ARRAY[1..ungGr05CylinderPosMaxNo] OF WORD;					(* Position cylinder status *)
	arlrAxisClampActPos					:ARRAY[1..ungGr05ClampMaxNo] OF LREAL;						(* Axis clamp actual position *)
	arlrAxisClampActVelo					:ARRAY[1..ungGr05ClampMaxNo] OF LREAL;						(* Axis clamp actual velocity *)
	arlrAxisClampActForce					:ARRAY[1..ungGr05ClampMaxNo] OF LREAL;						(* Axis clamp actual force *)
	unSawingStep						:UINT;						(* Current sawing step *)
END_STRUCT
END_TYPE

// ---- Data types/Machine/SEW/CIA402/ST_PLCTOSEWMOVIEDRIVEBCIA402.TcDUT
(* Communication structure from plc to drive *)

TYPE ST_PLCTOSEWMOVIEDRIVEBCIA402 :
STRUCT
	wPO1ControlWord			:WORD;
END_STRUCT
END_TYPE

// ---- Data types/Machine/SEW/CIA402/ST_SEWMOVIEDRIVEBCIA402TOPLC.TcDUT
(* Communikation structure from drive to plc *)

TYPE ST_SEWMOVIEDRIVEBCIA402TOPLC :
STRUCT
	wPO1StatusWord						:WORD;
	bAxisWeldingLimitMax 					:BOOL; 						(* DI1.5 Maximum limit of  axis welding / Endschalter Achse Schweißen maximal *)
	bAxisWeldingLimitMin 					:BOOL;						(* DI1.4 Minimum limit of  axis welding / Endschalter Achse Schweißen minimal *)
END_STRUCT
END_TYPE

// ---- Data types/Machine/SEW/CIA402/ST_SEWMOVIEDRIVEBCIA402_REF.TcDUT
TYPE ST_SEWMOVIEDRIVEBCIA402_REF : FB_SEWMOVIDRIVEBCIA402_REF;
END_TYPE

// ---- Data types/Machine/STOEBER/PS6A34/ST_STOEBER_PS6A34Status.TcDUT
(* Status of Stober PS6A34 *)

TYPE ST_STOEBER_PS6A34Status :
STRUCT
	bReady				:BOOL;			(* Stoeber PS6A34 ready / StoeberPS6A34 i.O. *)
	bNoOverload			:BOOL;			(* StoeberPS6A34 no overload  / StoeberPS6A34 nicht überlastet *)
	bGridPhaseOk		:BOOL;			(* StoeberPS6A34 no grid phase failure  / StoeberPS6A34 nicht Netzphasenausfall *)
END_STRUCT
END_TYPE

// ---- Data types/Machine/STOEBER/SDS/ST_BaseDeviceIn.TcDUT
TYPE ST_BaseDeviceIn :
STRUCT

	bEnabled					:BOOL;			(* The drive is ready for operation. *)
	bError						:BOOL;			(* The drive state is fault. *)
	bGroupError					:BOOL;			(* Group error: Maximum following error *)
	bQuickStop 					:BOOL;			(* Quick stop is queued/is being executed. *)
	bAxisActive					:BOOL;			(* Axis is active. *)
	bToggleBit 					:BOOL;			(* Handshake bit. *)

	(* Command Positioning *)
	stCommandPositioning			:ST_CommandPositioningFROMNC;

	(* Fast Referene Value  *)
	stFastRefereneValue			:ST_FastRefereneValueFROMNC;
END_STRUCT
END_TYPE

// ---- Data types/Machine/STOEBER/SDS/ST_BaseDeviceOut.TcDUT
TYPE ST_BaseDeviceOut :
STRUCT

	bEnable						:BOOL;			(* Enable controller *)
	bFaultReset					:BOOL;			(* Acknowledgment for faults of the device state machine. *)
	bQuickStop					:BOOL;			(* Brakes the motor *)
	bFeedEnablePlus				:BOOL;			(* Feed enable plus *)
	bFeedEnableMinus			:BOOL;			(* Feed enable minus *)
	bHomingSensor				:BOOL;			(* Referencing cam signal or homing sensor *)
	bToggleBit 					:BOOL;			(* Handshake bit. *)
	nTorqueLimit					:INT;			(* Value of torque limit (absolute value) *)

	(* Command Positioning *)
	stCommandPositioning			:ST_CommandPositioningFROMPLC;

	(* Fast Referene Value *)
	stFastRefereneValue			:ST_FastRefereneValueFROMPLC;

END_STRUCT
END_TYPE

// ---- Data types/Machine/STOEBER/SDS/ST_PLCTOSTOEBER.TcDUT
(* Communikation structure from plc to nc *)

TYPE ST_PLCTOSTOEBER :
STRUCT
	dnI34ReferencePosition				:DINT;
	dnI213TargetPosition					:DINT;
	nI230Override							:INT;
	nI215VeloFaktor						:INT;
	nD230NReferenceValueRelative		:INT;
	nC230TorqueLimit						:INT;
	wI210PosiControlWord					:WORD;
	wDummy1							:WORD;
	usnI216AccFaktor						:USINT;
	usnI217DccFaktor						:USINT;
	byA180DeviceControlByte				:BYTE;
	byI211MotionCommandByte			:BYTE;
END_STRUCT
END_TYPE

// ---- Data types/Machine/STOEBER/SDS/ST_STOEBERTOPLC.TcDUT
(* Communikation structure from nc to plc *)

TYPE ST_STOEBERTOPLC :
STRUCT
	dnI88Speed							:DINT;
	dnI203CurrentPosition					:DINT;
	nE90MMotor							:INT;
	nE100MMotor							:INT;
	unI200PosiStatusWord					:UINT;
	nD200SpeedReferenceValueStatusWord	:UINT;
	byE200DeviceStatusByte				:BYTE;
	byI201MotionStatusByte				:BYTE;
	byI90ErrorCode						:BYTE;
	byDummy1							:BYTE;
END_STRUCT
END_TYPE

// ---- Data types/Machine/STOEBER/SI6_SC6/CIA402/ST_CIA402In.TcDUT
TYPE ST_CIA402In :
STRUCT

	bReadyToSwitchOn 			:BOOL;			(* Ready to switch on. *)
	bSwitchedOn 					:BOOL;			(* Switched on. *)
	bEnabled 					:BOOL;			(* Operation enabled. *)
	bError  						:BOOL;			(* The drive state is fault. *)
	bVoltageEnabled 				:BOOL;			(* Voltage enabled. *)
	bQuickStop 					:BOOL;			(* Quick stop is queued/is being executed. *)
	bSwitchOnDisabled 			:BOOL;			(* Switch on disabled. *)
	bMessage 					:BOOL;			(* Message *)
	snDecimalDigits 				:SINT;			(* Number of positions after the decimal point for indication and entry of position reference values, speeds, accelerations *)

	(* Jog mode *)

	(* Position mode *)
	stPositionMode				:ST_PositionModeFromDrive;

	(* Velocity mode *)
	stVelocityMode				:ST_VelocityModeFromDrive;

	(* Torque mode *)
	stTorqueMode				:ST_TorqueModeFromDrive;

	(* Homing mode *)
	stHomingMode				:ST_HomingModeFromDrive;


	etModesOfOperation			:ET_ModesOfOperation;			(* Actual operating mode *)
																(*
																	-1: Jog
																	0: No mode assigned
																	1: Profile position mode
																	3: Profile velocity mode
																	4: Profile torque mode
																	6: Homing Mode
																	7: Interpolated position mode
																	8: Cyclic synchronous position mode
																	9: Cyclic synchronous velocity mode
																	10: Cyclic synchronous torque mode													
																*)
	dnActPosition					:DINT;			(* Actual position of the axis *)
	dnActVelocity					:DINT;			(* Actual velocity of the axis *)
	nActTorque 					:INT;			(* Actual torque/force of the axis *)
	dnActFollowingError			:DINT;			(* Actual lag *)

	bNegLimitSwitch				:BOOL;			(* Negative limit switch *)
	bPosLimitSwitch				:BOOL;			(* Positive limit switch *)
	bHomeSwitch 				:BOOL;			(* Reference switch *)

	dnActAdditionalPosition		:DINT;			(* Actual position of the master encoder *)


	snPLCOpenState				:SINT;
	snPLCOpenErrStopCause		:SINT;			(* Cause of a requested command being denied or cancelled by the motion core *)
	bPLCOpenError				:BOOL;			(* Motion core has denied or is cancelling the requested command  *)
	bPLCOpenDone				:BOOL;			(* The motion core has successfully ended the command to be executed  *)
	bPLCOpenAborted			:BOOL;			(* The motion core has aborted  *)

	bConstantVelocity				:BOOL;			(* Speed reached *)
	bAccelerating					:BOOL;			(* Accelerating  *)
	bDecelerating				:BOOL;			(* Decelerating  *)
	bNotMoving					:BOOL;			(* Actual speed is zero *)
	bReferenced					:BOOL;			(* Referenced *)

	dwDigitalInputs				:DWORD;

END_STRUCT
END_TYPE

// ---- Data types/Machine/STOEBER/SI6_SC6/CIA402/ST_CIA402Out.TcDUT
TYPE ST_CIA402Out :
STRUCT

	bSwitchOn 						:BOOL;			(* Switch on. *)
	bEnableVoltage					:BOOL;			(* Enable voltage *)
	bQuickStop						:BOOL;			(* Quick stop; 0 = request quick stop; 1 = do not request quick stop*)
	bEnableOperation					:BOOL;			(* Enable operation *)
	bFaultReset						:BOOL;			(* Fault reset 0, 1 = inactive; 0 -> 1 = active*)
	bHalt							:BOOL;			(* Prerequisite: Jog, Profile position, Profile velocity or Profile torque operating modes *)
	bOperatingModeSpecific			:BOOL;			(* Operating mode specific  *)
	bAxisSelectorBit0 					:BOOL;			(* Prerequisite: A63 = 2: Parameter  *)
	bAxisSelectorBit1 					:BOOL;			(* Prerequisite: A643 = 2: Parameter  *)
													(*
														00 bin = axis 1, 01 bin = axis 2, 10 bin = axis 3, 11 bin = axis 4
													*)
	bAxisDisable						:BOOL;			(* Prerequisite: A65 = 2: Parameter, 0 = do not disable axis; 1 = disable axis  *)
	bOpenBrake						:BOOL;			(* Prerequisite: F06 = 2: Parameter; 0 = brake control through device control (prerequisite: F92[0] = 0: Internal (automatic)) or 0 = engage brake (prerequisite: F92[0] = 1: External (plc)), 1 = open brake*)
	bSetReference					:BOOL;			(* Prerequisite: I111 = 2: Parameter, 0, 1 = inactive; 0 -> 1 = set reference without interrupting active movements; for controller-controlled operation, the controller must track the set position accordingly *)

	bFeedEnablePlus					:BOOL;			(* Feed enable plus *)
	bFeedEnableMinus				:BOOL;			(* Feed enable minus *)

	(* Jog mode *)
	stJogMode						:ST_JogModeFromPLC;

	(* Position mode *)
	stPositionMode					:ST_PositionModeFromPLC;

	(* Velocity mode *)
	stVelocityMode					:ST_VelocityModeFromPLC;

	(* Torque mode *)
	stTorqueMode					:ST_TorqueModeFromPLC;

	(* Homing mode *)
	stHomingMode					:ST_HomingModeFromPLC;


	etModesOfOperation				:ET_ModesOfOperation;			(* Set operating mode. *)
																	(*
																		-1: Jog
																		0: No mode assigned
																		1: Profile position mode
																		3: Profile velocity mode
																		4: Profile torque mode
																		6: Homing Mode
																		7: Interpolated position mode
																		8: Cyclic synchronous position mode
																		9: Cyclic synchronous velocity mode
																		10: Cyclic synchronous torque mode
																	*)

	nOverride						:INT;			(* Value of override 16384 = 100 %. *)
	unMaxTorque						:UINT;			(* Maximum permissible torque/force *)
	udnMaxAcceleration				:UDINT;			(* Maximum permissible acceleration in the Homing, Jog, Profile position and Profile velocity operating modes. *)
	udnMaxDeceleration				:UDINT;			(* Maximum permissible deceleration in the Homing, Jog, Profile position and Profile velocity operating modes. *)
	udnMaxJerk						:UDINT;			(* Maximum permitted jerk. *)
	dnSoftwarePosLimitMin				:DINT;			(* Positions of the software position limitation minimum *)
	dnSoftwarePosLimitMax			:DINT;			(* Positions of the software position limitation maximum *)

	dwDigitalOutputs 					:DWORD;

END_STRUCT
END_TYPE

// ---- Data types/Machine/STOEBER/SI6_SC6/CIA402/ST_PLCTOSTOEBERSI6SC6CIA402.TcDUT
(* Communikation structure from plc to drive *)

TYPE ST_PLCTOSTOEBERSI6SC6CIA402 :
STRUCT
	wA515Controlword					:WORD;
	snA541ModesOfOperation			:SINT;
	snDummy1						:SINT;
	dnA567TargetPosition				:DINT;
	dnA638TargetVelocity				:DINT;
	nA558TargetTorque 				:INT;
	unA559MaxTorque 				:UINT;
	udnA604MaxAcceleration			:UDINT;
	udnA605MaxDeceleration			:UDINT;
	udnA574Velocity					:UDINT;
	udnA576Acceleration				:UDINT;
	udnA577Deceleration				:UDINT;
	dnA569HomeOffset				:DINT;
	dnA570SoftwarePosLimitMin		:DINT;
	dnA570SoftwarePosLimitMax		:DINT;
	dwA637DigitalOutputs 				:DWORD;
END_STRUCT
END_TYPE

// ---- Data types/Machine/STOEBER/SI6_SC6/CIA402/ST_STOEBERSI6SC6CIA402TOPLC.TcDUT
(* Communikation structure from drive to plc *)

TYPE ST_STOEBERSI6SC6CIA402TOPLC :
STRUCT
	wA516Statusword						:WORD;
	snA542ModesOfOperationDisplay		:SINT;
	snDummy1							:SINT;
	dnA545PositionActualValue				:DINT;
	dnA553VelocityActualValue 			:DINT;
	nA564TorqueActualValue 				:INT;
	nDummy1							:INT;
	dnA632FollowingErrorActualeValue		:DINT;
	dnA620AdditionalPositionActualValue	:DINT;
	snI89PLCOpenState					:SINT;
	snI90PLCOpenErrStopCause			:SINT;
	wA67UserStatusword 					:WORD;
	dwA636DigitalInputs					:DWORD;
END_STRUCT
END_TYPE

// ---- Data types/Machine/STOEBER/SI6_SC6/CIA402/ST_STOEBERSI6SC6CIA402_REF.TcDUT
TYPE ST_STOEBERSI6SC6CIA402_REF : FB_STOEBERSI6SC6CIA402_REF;
END_TYPE

// ---- Data types/Machine/STOEBER/ST_STOEBER_AxisStatus.TcDUT
(* Status of Stober inverter *)

TYPE ST_STOEBER_AxisStatus :
STRUCT
	bEnabled					:BOOL;			(* Enabled = TRUE indicates that the inverter is enabled. *)
	bError						:BOOL;			(* Error = TRUE indicates that the inverter has error.*)
	bFastStopActive				:BOOL;			(* FastStopActive = TRUE indicates that the fast stop is active.*)
	bReadyToPos				:BOOL;			(* ReadyToPos = TRUE indicates that the inverter is ready to positioning.*)
	bLocalActive					:BOOL;			(* LocalActive = TRUE indicates that the local mode active.*)
	bJogActive					:BOOL;			(* JogActive = TRUE indicates that the jog mode active.*)
	bConstantVelocity               		:BOOL;			(* ConstantVelocity = TRUE indicates that the inverter is in velocity *)
	bAccelerating					:BOOL;			(* Drive is accelerating *)
	bDecelerating				:BOOL;			(* Drive is decelerating *)
	bInPosition					:BOOL;			(* InPosition = TRUE indicates that the inverter is in position.*)
	bInPositionWindow			:BOOL;			(* InPositionWindow = TRUE indicates that the inverter is in position window.*)
	bInReference					:BOOL;			(* InReference = TRUE indicates that the inverter is in reference.*)
	bStandStill					:BOOL;			(* StandStill = TRUE indicates that the inverter has stand still.*)
	bInSync						:BOOL;			(* InSync = TRUE indicates that the inverter in sync.*)
	bHoming						:BOOL;			(* Homing = TRUE indicates that the referencing is active.*)
	bCam1						:BOOL;			(* Cam1 = TRUE indicates that the cam 1 active.*)
	bSwitchPoint					:BOOL;			(* SwitchPoint = TRUE indicates that the switch point active.*)
	bDenied						:BOOL;			(* Denied = TRUE indicates that the command denied .*)
	bLimitSwitch					:BOOL;			(* LimitSwitch = TRUE indicates that the hard- oder software limit switch touched.*)
	nActMotionID					:INT;			(* ActMotionID = TRUE indicates that the actual motion ID.*)
	lrActPosition					:REAL;			(* ActPosition = TRUE indicates that the actual position.*)
END_STRUCT
END_TYPE

// ---- Data types/Machine/WeldingPhases/ET_WeldingDirection.TcDUT
TYPE ET_WeldingDirection :
(
	ET_WeldingDirection_eCurrent := 0,
	ET_WeldingDirection_ePositive := 1,
	ET_WeldingDirection_eNegative := -1
);
END_TYPE

// ---- Data types/Machine/WeldingPhases/Force/ST_BeadUp.TcDUT
TYPE ST_BeadUp :
STRUCT
	lrBeadUpForce						:LREAL;											(* BeadUp force [N] *)
	unBeadUpRamp						:UINT;											(* BeadUp ramp [s] *)
	unBeadUpTime						:UINT;											(* BeadUp time [s] *)
	lrVeloForceCtrlKp						:LREAL;											(* Velocity - force controller proportional band Kp *)
	lrVeloForceCtrlTi						:LREAL;											(* Velocity - force controller integral Ti *)
	lrVeloForceCtrlLimit					:LREAL;											(* Velocity - force controller limit  *)
END_STRUCT
END_TYPE

// ---- Data types/Machine/WeldingPhases/Force/ST_ForceProcess.TcDUT
TYPE ST_ForceProcess :
STRUCT
	lrProcessForce						:LREAL;											(* Process force [N] *)
	unProcessRamp						:UINT;											(* Process ramp [s] *)
	unProcessTime						:UINT;											(* Process time [s]  *)
	arunDuration							:ARRAY[1..2] OF UINT;								(* Duration [s] *)
	lrVeloForceCtrlKp						:LREAL;											(* Velocity - force controller proportional band Kp *)
	lrVeloForceCtrlTi						:LREAL;											(* Velocity - force controller integral Ti *)
	lrVeloForcePreCtrlVelo					:LREAL;											(* Feedforward velocity precontrol wieghting =  0..1 *)
	lrVeloForceCtrlLimit					:LREAL;											(* Velocity - force controller limit  *)
END_STRUCT
END_TYPE

// ---- Data types/Machine/WeldingPhases/Force/ST_ForceWelding.TcDUT
TYPE ST_ForceWelding :
STRUCT
	lrWeldingForce						:LREAL;											(* Welding force [N] *)
	unWeldingRamp						:UINT;											(* Welding ramp [s] *)
	unCoolDownTime						:UINT;											(* Cool down time [s]  *)
	arunCoolingTime						:ARRAY[1..2] OF UINT;								(* Cooling time *)
	lrVeloForceCtrlKp						:LREAL;											(* Velocity - force controller proportional band Kp *)
	lrVeloForceCtrlTi						:LREAL;											(* Velocity - force controller integral Ti *)
	lrVeloForcePreCtrlVelo					:LREAL;											(* Feedforward velocity precontrol wieghting =  0..1 *)
	lrVeloForceCtrlLimit					:LREAL;											(* Velocity - force controller limit  *)
END_STRUCT
END_TYPE

// ---- Data types/Machine/WeldingPhases/Force/ST_HeatUp.TcDUT
TYPE ST_HeatUp :
STRUCT
	lrHeatUpForce						:LREAL;											(* HeatUp force [N] *)
	unHeatUpRamp						:UINT;											(* HeatUp ramp [s] *)
	unHeatUpTime						:UINT;											(* HeatUp time [s] *)
	lrVeloForceCtrlKp						:LREAL;											(* Velocity - force controller proportional band Kp *)
	lrVeloForceCtrlTi						:LREAL;											(* Velocity - force controller integral Ti *)
	lrVeloForceCtrlLimit					:LREAL;											(* Velocity - force controller limit  *)
END_STRUCT
END_TYPE

// ---- Data types/Machine/WeldingPhases/Force/ST_PreHeat.TcDUT
TYPE ST_PreHeat :
STRUCT
	lrPreHeatForce						:LREAL;											(* PreHeat force [N] *)
	unPreHeatRamp						:UINT;											(* PreHeat ramp [s] *)
	unPreHeatTime						:UINT;											(* PreHeat time [s] *)
	lrVeloForceCtrlKp						:LREAL;											(* Velocity - force controller proportional band Kp *)
	lrVeloForceCtrlTi						:LREAL;											(* Velocity - force controller integral Ti *)
	lrVeloForcePreCtrlVelo					:LREAL;											(* Feedforward velocity precontrol wieghting =  0..1 *)
	lrVeloForceCtrlLimit					:LREAL;											(* Velocity - force controller limit  *)
END_STRUCT
END_TYPE

// ---- Data types/Machine/WeldingPhases/Force/ST_WeldingPhases.TcDUT
TYPE ST_WeldingPhases :
STRUCT
	stPreHeat							:ST_PreHeat;
	stBeadUp							:ST_BeadUp;
	stHeatUp							:ST_HeatUp;
	unChangeoverTime					:UINT;											(* Changeover time [s] *)
	stWelding							:ST_ForceProcess;
END_STRUCT
END_TYPE

// ---- Data types/Machine/WeldingPhases/Position/ST_PositionProcess.TcDUT
TYPE ST_PositionProcess :
STRUCT
	lrProcessPosition						:LREAL;											(* Process position [mm] *)
	unProcessVelo						:UINT;											(* Process force [%] *)
	unProcessRamp						:UINT;											(* Process ramp [s] *)
	unProcessTime						:UINT;											(* Process time [s]  *)
	arunDuration							:ARRAY[1..2] OF UINT;								(* Duration [s] *)
END_STRUCT
END_TYPE

// ---- Data types/Machine/WeldingPhases/Position/ST_PositionWelding.TcDUT
TYPE ST_PositionWelding :
STRUCT
	lrWeldingPosition						:LREAL;											(* Welding position [mm] *)
	unWeldingVelo						:UINT;											(* Welding force [%] *)
	unWeldingRamp						:UINT;											(* Welding ramp [s] *)
	unCoolDownTime						:UINT;											(* Cool down time [s]  *)
	arunCoolingTime						:ARRAY[1..2] OF UINT;								(* Cooling time *)
END_STRUCT
END_TYPE

// ---- Data types/Machine/WeldingPhases/ST_WeldingStatus.TcDUT
TYPE ST_WeldingStatus :
STRUCT
	lrStartWelding				:LREAL;
	lrEndWelding					:LREAL;
	lrDistanceWelding				:LREAL;
END_STRUCT
END_TYPE

// ---- Data types/Objects/Axis/ExternelMC/ET_JogMode.TcDUT
TYPE ET_JogMode :
(
	ET_JogMode_MC_JOGMODE_STANDARD,
	ET_JogMode_MC_JOGMODE_INCHING
);
END_TYPE

// ---- Data types/Objects/Axis/ExternelMC/ET_MC_Direction.TcDUT
TYPE ET_MC_Direction :
(
	ET_MC_Direction_eCurrent := 0,
	ET_MC_Direction_ePositive := 1,
	ET_MC_Direction_eNegative := -1
);
END_TYPE

// ---- Data types/Objects/Axis/ExternelMC/ET_MC_States.TcDUT
TYPE ET_MC_States :
(
	ET_MC_States_eInit := 100,
	ET_MC_States_eReset,
	ET_MC_States_eRunning,
	ET_MC_States_eWaiting,
	ET_MC_States_eAbort,
	ET_MC_States_eDone,
	ET_MC_States_eError,
	ET_MC_States_eNotExecute
);
END_TYPE

// ---- Data types/Objects/Axis/ExternelMC/SDS/ST_CommandPositioningFROMNC.TcDUT
TYPE ST_CommandPositioningFROMNC :
STRUCT
	(* Command Positioning *)
	bConstantVelocity				:BOOL;			(* Constant speed reached. *)
	bHomed						:BOOL;			(* Axis is referenced. *)
	bPositionReached			:BOOL;			(* Window around target position reached for the first time. *)
	bPositionWinReached			:BOOL;			(* Actual position is located in the position window. *)
	bNotMoving					:BOOL;			(* Axis is logically stationary. *)
	bDenied						:BOOL;			(* Indicates that the command denied .*)
	bCoupled 					:BOOL;			(* Axis coupling state *)
	dnActPosition					:DINT;			(* Value of current (actual) position *)
	dnActVelocity					:DINT;			(* Value of current (actual) velocity *)
	nActEngineTorque			:INT;			(* Indication of the current motor torque in Nm *)
	rDecimalDigits 				:REAL;			(* Number of positions after the decimal point for indication and entry of position reference values, speeds, accelerations *)
	udnScalingDenom				:UDINT := 1;	  	(* Effective distance per rev. Denominator [INC] *)
	lrScalingNum					:LREAL;			(* Effective distance per rev. Numerator [technical units]: The factor indicates the distance per one increment of position control.*)
	bLimitMaxExceeded			:BOOL;			(* Position limit switch maximum is exceeded *)
	bLimitMinExceeded			:BOOL;			(* Position limit switch minimum is exceeded *)

	byPLCOpenState				:BYTE;			(* Supplies information on the reaction of the axis during operation on a fieldbus. *)
	bPLCOpenStandstill			:BOOL;			(* PLCopen state Standstill. *)
	bPLCOpenCmdAborted		:BOOL;			(* Positioning command denied/aborted. TRUE means that the last positioning job was aborted. *)
	bPLCOpenCmdDone			:BOOL;			(* TRUE means that the command was executed successfully. *)
	byPLCOpenErrorCode			:BYTE;			(* When the PLCOpen state is ErrorStop. *)

END_STRUCT
END_TYPE

// ---- Data types/Objects/Axis/ExternelMC/SDS/ST_CommandPositioningFROMPLC.TcDUT
TYPE ST_CommandPositioningFROMPLC :
STRUCT
	(* Command Positioning *)
	nOverride					:INT;			(* Value of override 16384 = 100 %. *)
	nVeloFactor					:INT;			(* Value of the velocity 16384 = 100 %. *)
	usnAccFactor					:USINT;			(* Value of the acceleration (always positive) 255 = 100% *)
	usnDccFaktor					:USINT;			(* Value of the deceleration (always positive) 255 = 100% *)
	usnJerkFaktor				:USINT;			(* Value of the jersk (always positive) 255 = 100% *)
	dnTargetPosition				:DINT;			(* Value of target position *)
	dnReferencePosition			:DINT;			(* Value which is loaded as the actual position in the reference point. *)
	bTipEnable					:BOOL;			(* Activates tipping mode. *)
	bTipPlus						:BOOL;			(* Tip mode in positive direction. *)
	bTipMinus					:BOOL;			(* Tip mode in negative direction. *)

	byPLCOpenCmd				:BYTE;			(* Global parameter for specification of the command to be executed via fieldbus. *)
	bPLCOpenCmdExe			:BOOL;			(* With a rising edge, the command in Motion Command is executed. *)

END_STRUCT
END_TYPE

// ---- Data types/Objects/Axis/ExternelMC/SDS/ST_DRIVE_REF.TcDUT
TYPE ST_DRIVE_REF : FB_STOEBERSDS_Drive_REF;
END_TYPE

// ---- Data types/Objects/Axis/ExternelMC/SDS/ST_FastRefereneValueFROMNC.TcDUT
TYPE ST_FastRefereneValueFROMNC :
STRUCT
	(* Fast Referene Value *)
	bStandstill					:BOOL;			(* Standstill. *)
	bVeloReached				:BOOL;			(* Reference value reached *)
	nMotorSpeed					:INT;			(* Current motor speed *)
END_STRUCT
END_TYPE

// ---- Data types/Objects/Axis/ExternelMC/SDS/ST_FastRefereneValueFROMPLC.TcDUT
TYPE ST_FastRefereneValueFROMPLC :
STRUCT
	(* Fast Referene Value *)
	nOverride					:INT;			(* Value of override 16384 = 100 %. *)
	nSpeed						:INT;			(* Relative speed reference value *)
	bHWLimitMax					:BOOL;			(* Hardware limit switch maximum end of range *)
	bHWLimitMin					:BOOL;			(* Hardware limit switch minimum end of range *)
END_STRUCT
END_TYPE

// ---- Data types/Objects/Axis/ExternelMC/SI6/ET_ModesOfOperation.TcDUT
TYPE ET_ModesOfOperation :
(
	ET_ModesOfOperation_Jog := -1,							(* -1: Jog *)
	ET_ModesOfOperation_None := 0,							(* 0: No mode assigned *)
	ET_ModesOfOperation_ProfilePosition := 1,					(* 1: Profile position mode *)
	ET_ModesOfOperation_Velocity := 2,							(* 2: Profile velocity mode *)
	ET_ModesOfOperation_ProfileVelocity := 3,					(* 3: Profile velocity mode *)
	ET_ModesOfOperation_ProfileTorque := 4,					(* 4: Profile torque mode *)
	ET_ModesOfOperation_Inactive := 5,							(* 5: Inactive *)
	ET_ModesOfOperation_Homing := 6,							(* 6: Homing Mode *)
	ET_ModesOfOperation_InterpolatedPosition := 7,				(* 7: Interpolated position mode *)
	ET_ModesOfOperation_CyclicSynchroPosition := 8,				(* 8: Cyclic synchronous position mode *)
	ET_ModesOfOperation_CyclicSynchroVelocity := 9,				(* 9: Cyclic synchronous velocity mode *)
	ET_ModesOfOperation_CyclicSynchroTorque := 10				(* 10: Cyclic synchronous torque mode *)
);
END_TYPE

// ---- Data types/Objects/Axis/ExternelMC/SI6/ST_DRIVESI6SC6CIA402_REF.TcDUT
TYPE ST_DRIVESI6SC6CIA402_REF : FB_STOEBERSI6SC6CIA402_REF;
END_TYPE

// ---- Data types/Objects/Axis/ExternelMC/SI6/ST_HomingModeFromDrive.TcDUT
TYPE ST_HomingModeFromDrive :
STRUCT
	bHomeReached				:BOOL;			(* Referencing ended  *)
	bHomingAttained				:BOOL;			(* Reference set *)
	bHomingError				:BOOL;			(* Referencing error *)
												(*
													000 bin = referencing active; 
													001 bin = referencing canceled or not started; 
													010 bin = reference set, referencing not yet complete; 
													011 bin = referencing ended successfully; 
													100 bin = referencing error, velocity is not zero; 
													110 bin = referencing error, velocity is zero
												*)
END_STRUCT
END_TYPE

// ---- Data types/Objects/Axis/ExternelMC/SI6/ST_HomingModeFromPLC.TcDUT
TYPE ST_HomingModeFromPLC :
STRUCT
	bHomingOperationStart			:BOOL;			(* Start referencing 0, 1 = inactive; 0 -> 1 = active *)
	snHomingMethod					:SINT;			(* Set reference method for the Homing operating mode. *)
	dnHomeOffset					:DINT;			(* Reference position of the axis in the Homing operating mode and for the Set reference function *)
END_STRUCT
END_TYPE

// ---- Data types/Objects/Axis/ExternelMC/SI6/ST_JogModeFromPLC.TcDUT
TYPE ST_JogModeFromPLC :
STRUCT
	bJogPositive					:BOOL;			(* 0 = inactive; 1 = active *)
	bJogNegative				:BOOL;			(* 0 = inactive; 1 = active *)
	dnJogStep					:DINT;			(* Jog step *)
	lrVelocity						:LREAL;			(* Jog velocity *)
	lrAcceleration					:LREAL;			(* Acceleration in the Jog. *)
	lrDeceleration				:LREAL;			(* Deceleration in the Jog. *)
	lrJerk						:LREAL;			(* Jerk  in the Jog. *)
END_STRUCT
END_TYPE

// ---- Data types/Objects/Axis/ExternelMC/SI6/ST_PositionModeFromDrive.TcDUT
TYPE ST_PositionModeFromDrive :
STRUCT
	bPositionReached			:BOOL;			(* Set position reached, data source: I180; prerequisite: halt inactive = A515, bit 8 = 0
												    Velocity is zero; data source: I199; prerequisite: halt inactive = A515, bit 8 = 1 *)
	bSetpointAck					:BOOL;			(* Target position accepted from motion core *)
	bFollowingError				:BOOL;			(* Following error *)
END_STRUCT
END_TYPE

// ---- Data types/Objects/Axis/ExternelMC/SI6/ST_PositionModeFromPLC.TcDUT
TYPE ST_PositionModeFromPLC :
STRUCT
	(* Command Positioning *)
	dnTargetPosition					:DINT;			(* Target position of the Profile position operating mode and set position of the Cyclic synchronous position operating mode. *)
	bNewSetpoint					:BOOL;			(* New setpoint (apply the new target position and start the movement) 0, 1 = inactive; 0 -> 1 = active *)
	bChangeSetImmediately			:BOOL;			(* 0 = apply new target position with bit 4 if no movement is active (prerequisite: I199 = 1: Active); 1 = apply new target position always with bit 4; a movement that is still active is interrupted *)
	bAbsRel							:BOOL;			(* Absolute target position/relative distance; 0 = Target position is an absolute position; 1 = Target position is a distance relative to the last target position A567 (prerequisite: A621 = X to X00 bin) or 1 = Target position is a distance relative to the current actual position A545 (prerequisite: A621 = X to X10 bin) *)
	udnVelocity						:UDINT;			(* Velocity for profile. *)
	udnAcceleration					:UDINT;			(* Acceleration for profile. *)
	udnDeceleration					:UDINT;			(* Deceleration for profile. *)
	udnJerk							:UDINT;			(* Jerk  for profile. *)
END_STRUCT
END_TYPE

// ---- Data types/Objects/Axis/ExternelMC/SI6/ST_TorqueModeFromDrive.TcDUT
TYPE ST_TorqueModeFromDrive :
STRUCT
	bTorqueReached				:BOOL;			(* Set force / set torque reached; difference in the amount of effective set force / set torque and actual force / actual torque greater than torque / force window, data source: A558, A564, G900  *)
END_STRUCT
END_TYPE

// ---- Data types/Objects/Axis/ExternelMC/SI6/ST_TorqueModeFromPLC.TcDUT
TYPE ST_TorqueModeFromPLC :
STRUCT
	nTargetTorque 					:INT;			(* Set torque/force in the Profile torque operating mode *)
END_STRUCT
END_TYPE

// ---- Data types/Objects/Axis/ExternelMC/SI6/ST_VelocityModeFromDrive.TcDUT
TYPE ST_VelocityModeFromDrive :
STRUCT
	bVelocityReached			:BOOL;			(* set velocity reached; data source: I85; prerequisite: halt inactive = A515, bit 8 = 0
												    Velocity is zero; data source: I199; prerequisite: halt inactive = A515, bit 8 = 1 *)
	bVelocityZero				:BOOL;			(* Velocity is zero; data source I199 *)
	bMaxSlippageError			:BOOL;			(* Difference in the amount of the effective set and actual velocity greater than velocity window, data source: I426, I88, C40 *)
END_STRUCT
END_TYPE

// ---- Data types/Objects/Axis/ExternelMC/SI6/ST_VelocityModeFromPLC.TcDUT
TYPE ST_VelocityModeFromPLC :
STRUCT
	(* Command velocity *)
	dnTargetVelocity				:DINT;			(* Target velocity for Profile velocity operating mode. *)
	udnAcceleration				:UDINT;			(* Acceleration for profile. *)
	udnDeceleration				:UDINT;			(* Deceleration for profile. *)
	udnJerk						:UDINT;			(* Jerk  for profile. *)
END_STRUCT
END_TYPE

// ---- Data types/Objects/Axis/ExternelMC/ST_AXIS_REF.TcDUT
TYPE ST_AXIS_REF :
STRUCT
	sAdsAddr			:STRING(23);			(* AmsNetId of the EtherCAT master device.*)
	unSlaveAddr			:UINT;				(* Address of the slave device.*)
	bLockPDO			:BOOL;
	bCmdInterrupted		:BOOL;
	bHWLimitMax			:BOOL;
	bHWLimitMin			:BOOL;
	bSWLimitMax			:BOOL;
	bSWLimitMin			:BOOL;
	stNcToPlc			:ST_NCTOPLC;
	stPlcToNc			:ST_PLCTONC;
	stAxisStatus			:ST_STOEBER_AxisStatus;
	fbReadStatusSDS		:FB_STOEBERSDS_ReadStatus;
	fbReadStatusSI6		:FB_STOEBERSI6_ReadStatus;
END_STRUCT
END_TYPE

// ---- Data types/Objects/Axis/ExternelMC/ST_NCTOPLC.TcDUT
TYPE ST_NCTOPLC :
STRUCT
	(* SDS *)
	stBaseDevice				:ST_BaseDeviceIn;

	(* SD6/SC6/SI6 *)
	stCIA402						:ST_CIA402In;

END_STRUCT
END_TYPE

// ---- Data types/Objects/Axis/ExternelMC/ST_PLCTONC.TcDUT
TYPE ST_PLCTONC :
STRUCT
	(* SDS *)
	stBaseDevice				:ST_BaseDeviceOut;

	(* SD6/SC6/SI6 *)
	stCIA402						:ST_CIA402Out;



(*



	dnReferencePosition			:DINT;			(* Value which is loaded as the actual position in the reference point. *)

*)
END_STRUCT
END_TYPE

// ---- Data types/Objects/Axis/InternalMC/Controller/ET_MC_ControllerMode.TcDUT
TYPE ET_MC_ControllerMode :
(
	ET_MC_ControllerMode_eCMUndefined,
	ET_MC_ControllerMode_eCMTorque,
	ET_MC_ControllerMode_eCMVelocity,
	ET_MC_ControllerMode_eCMPosition,
	ET_MC_ControllerMode_eCMCurrent
	
);
END_TYPE

// ---- Data types/Objects/Axis/InternalMC/Controller/ST_VeloControllerConfig.TcDUT
TYPE ST_VeloControllerConfig :
STRUCT

	lrKp							:LREAL := 0.005;					(* Tuning parameter, proportional gain *)
	lrTi							:LREAL := 1000000;				(* Tuning parameter, time of integral *)
	lrTd							:LREAL := 0.0;						(* Tuning parameter, time of differential *)
	lrPreCtrlVelo					:LREAL := 0.01; 					(* Feedforward velocity precontrol wieghting =  0..1 *)
	lrVeloKpFilter					:LREAL := 1.0;						(* Velocity filter - proportional gain *)
	tVeloT1Filter					:TIME := t#100ms;					(* Velocity filter - time constant *)
	tDeadTime					:TIME := t#200ms;					(* Dead time *)
	lrDeltaMax					:LREAL := 100.0;					(* Maximum difference between two actual position values *)
	lrVeloMin					:LREAL := -100.0;					(* Velocity limit minimum [technical units / sec] *)
	lrVeloMax					:LREAL := 100.0;					(* Velocity limit maximum [technical units / sec] *)
	lrDeadZone					:LREAL := 10.0;					(* Dead zone *)

END_STRUCT
END_TYPE

// ---- Data types/Objects/Axis/InternalMC/Drive/ST_DriveConfig.TcDUT
TYPE ST_DriveConfig :
STRUCT
	
	bRealDrive					:BOOL := TRUE; 				(* Encoder ID number *) 

END_STRUCT
END_TYPE

// ---- Data types/Objects/Axis/InternalMC/Encoder/ST_EncoderConfig.TcDUT
TYPE ST_EncoderConfig :
STRUCT
	
